(* IEC 61131-3 sources: daoli-st-library/DL_Device (part 31) *)

(* ---- FB_DL_SlurryLevelBank.st ---- *)
(*
  FB_DL_SlurryLevelBank  —  多罐浆料液位开关组（fail-safe 方向解释 / 质量字仲裁 / 开关相反归因）/ Slurry level switch bank
  分类 Category : DL_Device
  码位 Code     : 16#03_2_0E
  版本 Version  : 1.0.0
  来源 Source   : t2-8-isa182 — IEC 61131-3 标准语义的道莅防御性实现
  溯源 Origin   : ISA-18.2 报警管理公开语义借鉴（报警与故障分离、状态归因），clean-room 实现，未复制源码行
  功能 Function : 1) 逐罐读取高位/低位点式开关、质量字（0~3，0 = OK）与组态 fail-safe 方向；
                  2) 按 fail-safe 方向解释「液位 vs 断线」：LOW 型（eLow）断线时读数表现为高位，
                     HIGH 型（eHigh）断线时读数表现为低位——两类方向各自反推，绝不套用同一公式；
                  3) 质量字非 OK 判 abSensorFault，并以**安全侧**值参与联锁（保守取值：保护泵的取「低」，
                     保护溢流的取「高」，即一律认报警成立），信息级 011E 记录替代生效；
                  4) 同一罐高低位同时为真判「开关相反」故障 022E（3 罐 × 2 型共 6 组向量逐条推演，见验收向量）；
                  5) 输出严格区分「越限（工艺）」与「传感器故障（仪表）」两类：越限只置 abLevelAlarm 与信息级 010E，
                     传感器故障置 abSensorFault 与故障级 021E 并置 bError（R190 归因唯一）。
  边界 Boundary : ① uBankSize = 0 或 > DL_BANK_MAX 判组态错 020E，**直接返回不进入循环**（防数组越界，R28-2）；
                     高位/低位/质量字/方向四个数组声明长度一律 DL_BANK_MAX，长度不等在编译期即被拦截，
                     运行期再以 uBankSize 做上界闸（双保险）；
                  ② 质量字不在 0~3 域内判组态错（质量字编码越界，无法解释），不按 OK 处理；
                  ③ fail-safe 方向枚举落 ELSE（非法方向）按「最保守」处理：高低两位都认报警，并置 020E；
                  ④ 解除式自证：_bFault 清除 = rtReset.Q（引脚可满足）；022E 另可由「该罐高低位不再同时为真」
                     按码专清（R188 可达清除边，不依赖人工复位掩盖真实接线错误）；
                  ⑤ nFaultCount 为 INT，逐罐故障计数后钳制到 DL_BANK_MAX（不溢出、不回绕）；
                  ⑥ 越限（010E）为信息级，**永不置 bError**（R187③ / R45 配对纪律）。
  依赖 Depends  : 仅 Standard.library（TON / R_TRIG / ABS / MIN / MAX），零外部组件依赖
  同拍双窗配比  : tQualityDb（质量字去抖）与心跳窗 DL_HEART_WINDOW 不同源；配比约束
                  tQualityDb <= DL_HEART_WINDOW，保证去抖窗内至少一次判活（R100）

  码表 Error codes（本件格 03_2_0E，子码步进 +0x10）:
    16#0003_020E 故障级：组态非法（uBankSize = 0 或越上限 / 质量字越 0~3 域 / fail-safe 方向非法）
    16#0003_021E 故障级：传感器故障（质量字非 OK，已用安全侧值参与联锁）
    16#0003_022E 故障级：开关相反（同一罐高低位同时为真，接线或组态错误）
    16#0003_023E 故障级：状态机落 ELSE 兜底（非法相位 ID）
    16#0003_010E 信息级：液位越限（工艺告警，不置 bError）
    16#0003_011E 信息级：断线安全侧替代已生效（保守取值，不置 bError）

  修订历史 Revision :
    2026-11-18  v1.0.0  R37 首版
*)

TYPE E_DL_FailSafeDir :
(
    eLow  := 0,   // 低液位型：液位低时开关动作；断线时读数浮为「高位」/ Low-level type, a broken wire reads as high
    eHigh := 10   // 高液位型：液位高时开关动作；断线时读数浮为「低位」/ High-level type, a broken wire reads as low
);
END_TYPE

TYPE E_DL_LevelBankState :
(
    eIdle  := 0,   // 空闲：未使能，输出全部复位 / Idle, all outputs cleared while disabled
    eRun   := 10,  // 运行：逐罐评估 / Running, per-tank evaluation
    eFault := 90   // 故障：组态非法锁定 / Fault, illegal configuration latched
);
END_TYPE

FUNCTION_BLOCK FB_DL_SlurryLevelBank
VAR_INPUT
    bEnable        : BOOL := FALSE;                       // 总使能，FALSE 时输出全复位 / Master enable, low level clears the outputs
    bReset         : BOOL := FALSE;                       // 复位，上升沿清故障锁存 / Reset, rising edge clears the latch
    uBankSize      : UINT := 3;                           // 罐组实际罐数 [个]，域 1~DL_BANK_MAX / Number of tanks in use
    abLevelHigh    : ARRAY[0..7] OF BOOL;                 // 高位开关原始输入 [BOOL/罐] / Raw high-level switch inputs
    abLevelLow     : ARRAY[0..7] OF BOOL;                 // 低位开关原始输入 [BOOL/罐] / Raw low-level switch inputs
    anSensorQuality : ARRAY[0..7] OF INT;                 // 传感器质量字 [0~3，0 = OK] / Sensor quality word, zero means OK
    aeFailSafeDir  : ARRAY[0..7] OF E_DL_FailSafeDir;     // 每罐 fail-safe 方向组态 [枚举/罐] / Per-tank fail-safe direction
    tQualityDb     : TIME := T#500MS;                     // 质量字去抖窗 [ms]，域 > 0 / Quality debounce window [ms]
END_VAR
VAR_OUTPUT
    abLevelAlarm   : ARRAY[0..7] OF BOOL;                 // 逐罐液位越限报警 [BOOL/罐] / Per-tank level alarm
    abSensorFault  : ARRAY[0..7] OF BOOL;                 // 逐罐传感器故障 [BOOL/罐] / Per-tank sensor fault
    nFaultCount    : INT;                                 // 故障罐数 [个] / Number of faulty tanks
    bBankAlarm     : BOOL;                                // 罐组总报警（越限或故障任一）/ Bank aggregate alarm
    bValid         : BOOL;                                // 判据可用标志 / Criteria usable
    bError         : BOOL;                                // 故障标志，派生自锁存 / Fault flag derived from the latch
    nErrId         : UDINT;                               // 事件码，0 = 无事件 / Event code, 0 = no event
    eStateOut      : E_DL_LevelBankState;                 // 状态出口，段尾单点映射 / State outlet, mapped at the tail
END_VAR
VAR
    tonQuality   : TON;                                   // 质量故障去抖窗，每拍无条件调用 / Quality fault debounce, called unconditionally
    tonHeart     : TON;                                   // 周期心跳窗，自复位 / Periodic heartbeat window, self-resetting
    rtReset      : R_TRIG;                                // 复位上升沿 / Reset rising edge
    _eState      : E_DL_LevelBankState := E_DL_LevelBankState.eIdle;  // 内部相位（CASE 唯一写入目标）/ Internal phase
    _uFault      : UDINT;                                 // 故障码锁存 / Latched fault code
    _uInfo       : UDINT;                                 // 信息码，每拍重算 / Information code, recomputed per scan
    _bFault      : BOOL;                                  // 故障锁存位 / Latched fault bit
    _bCfgBad     : BOOL;                                  // 组态非法聚合 / Configuration invalid aggregate
    _bAnySensFault : BOOL;                                // 任一罐传感器故障 / Any sensor fault present
    _bAnyOpposite  : BOOL;                                // 任一罐高低位相反 / Any opposite-switch condition
    _bAnyLevelAlarm : BOOL;                               // 任一罐液位越限 / Any level alarm present
    _bSafeSubst  : BOOL;                                  // 本拍发生安全侧替代 / A safe-side substitution happened
    _bOppClear   : BOOL;                                  // 相反故障已全部消失 / All opposite conditions cleared
    _bHeartBrk   : BOOL := TRUE;                          // 心跳窗断输入一拍 / One-scan heartbeat break
    _bQualBrk    : BOOL := TRUE;                          // 质量去抖断输入一拍 / One-scan quality break
    _nIdx        : INT;                                   // 循环索引 [索引] / Loop index
    _nFaultAcc   : INT;                                   // 故障罐数保持量 [个] / Held faulty-tank count
    _bHighEff    : BOOL;                                  // 高位开关的解释后值（含安全侧替代）/ Effective high-level value
    _bLowEff     : BOOL;                                  // 低位开关的解释后值（含安全侧替代）/ Effective low-level value
    _bOpposite   : BOOL;                                  // 本罐高低位同时为真 / Both switches true in this tank
    _bQualBad    : BOOL;                                  // 本罐质量字非 OK / Quality word not OK in this tank
    _bDirBad     : BOOL;                                  // 本罐方向枚举非法 / Illegal direction enumeration in this tank
END_VAR
VAR CONSTANT
    DL_BANK_MAX   : INT := 8;          // 数组声明长度 [个]，四数组同长 / Declared array length, identical for all four arrays
    DL_QUAL_MAX   : INT := 3;          // 质量字最大值 [编码] / Maximum quality code
    DL_HEART_WINDOW : TIME := T#2S;    // 心跳观察窗 [ms]，自复位节拍 / Heartbeat window, self-resetting
END_VAR

(* —— 段 0：定时器与边缘检测无条件周期刷新（R182：调用语句不得置于 IF / CASE / FOR 内） —— *)
rtReset(CLK := bReset);                                          // 复位上升沿，每拍必调
tonHeart(IN := (NOT tonHeart.Q) AND (NOT _bHeartBrk), PT := DL_HEART_WINDOW);  // 心跳窗自复位
_bHeartBrk := FALSE;                                             // 断输入拍在调用后自清
tonQuality(IN := (_eState = E_DL_LevelBankState.eRun) AND _bAnySensFault AND (NOT _bQualBrk),
           PT := tQualityDb);                                    // 质量故障去抖（表达式入参）
_bQualBrk := FALSE;                                              // 断输入拍在调用后自清

(* —— 段 1：单拍量预清零（数组输出与保持量不入清单，R187①） —— *)
_uInfo        := 16#0000_0000;   // 信息码每拍重算
bError        := FALSE;          // 故障出口每拍重算，段 6 由锁存派生
bValid        := FALSE;          // 可用标志缺省 FALSE
bBankAlarm    := FALSE;          // 罐组总报警缺省 FALSE
_bCfgBad      := FALSE;          // 组态非法预清零
_bAnySensFault := FALSE;         // 传感器故障聚合预清零
_bAnyOpposite := FALSE;          // 相反故障聚合预清零
_bAnyLevelAlarm := FALSE;        // 越限聚合预清零
_bSafeSubst   := FALSE;          // 安全侧替代标志预清零
_bOppClear    := TRUE;           // 相反故障清空判定初值（循环内遇相反即置 FALSE）
_bDirBad      := FALSE;          // 方向非法预清零

(* —— 段 2：复位沿清锁存 + 按码专清（R188 双路径） —— *)
IF rtReset.Q THEN
    _bFault     := FALSE;            // 复位沿清锁存位
    _uFault     := 16#0000_0000;     // 复位沿清锁存码
    _nFaultAcc  := 0;                // 复位沿清故障罐数（重新统计）
END_IF

(* —— 段 3：组态域闸（循环之前完成，越界即返回不进入循环，R28-2） —— *)
IF (uBankSize = 0) OR (uBankSize > INT_TO_UINT(DL_BANK_MAX)) THEN
    _bCfgBad := TRUE;                // 罐数越界：0 或超数组声明长度
END_IF
IF TIME_TO_DINT(tQualityDb) <= 0 THEN
    _bCfgBad := TRUE;                // 去抖窗非法
END_IF
IF _bCfgBad THEN
    _uFault := 16#0003_020E;         // 故障级：组态非法
    _bFault := TRUE;                 // 锁存位置位（复位沿可清）
    bError  := TRUE;                 // 故障标志置位（R45 配对）
    _eState := E_DL_LevelBankState.eFault;  // 进故障相（不进入循环）
END_IF

(* —— 段 4：逐罐评估（仅运行相且组态合法时进入；循环上界由 uBankSize 钳制） —— *)
IF bEnable AND (_eState <> E_DL_LevelBankState.eFault) AND (NOT _bCfgBad) THEN
    _nFaultAcc := 0;                          // 故障罐数每拍重算（输出量，非台账）
    FOR _nIdx := 0 TO (UINT_TO_INT(uBankSize) - 1) DO
        (* 4.1 本罐假设值初始化：有效值先取原始值，随后按质量与方向修正 *)
        _bHighEff := abLevelHigh[_nIdx];       // 高位原始读数 [BOOL]
        _bLowEff  := abLevelLow[_nIdx];        // 低位原始读数 [BOOL]
        _bQualBad := (anSensorQuality[_nIdx] < 0) OR (anSensorQuality[_nIdx] > DL_QUAL_MAX) OR
                     (anSensorQuality[_nIdx] <> 0);            // 质量字非 OK（含越域：无法解释即判坏）
        IF (anSensorQuality[_nIdx] < 0) OR (anSensorQuality[_nIdx] > DL_QUAL_MAX) THEN
            _bCfgBad := TRUE;                  // 质量字越 0~3 域：组态/采集链错误
            _uFault := 16#0003_020E;           // 故障级：组态非法
            _bFault := TRUE;                   // 锁存
            bError  := TRUE;                   // 故障标志置位（R45 配对）
        END_IF
        IF _bQualBad THEN
            _bAnySensFault := TRUE;            // 传感器故障聚合
            abSensorFault[_nIdx] := TRUE;      // 逐罐故障输出
            _bSafeSubst := TRUE;               // 发生安全侧替代
            (* 4.2 fail-safe 方向解释：断线时 LOW 型读成「高位」，HIGH 型读成「低位」——
                   保守取值即两者都按「报警成立」处理（低液位保护泵、高液位保护溢流） *)
            IF aeFailSafeDir[_nIdx] = E_DL_FailSafeDir.eLow THEN
                _bHighEff := FALSE;            // LOW 型断线：原始高位读数是浮空假象，不予采信
                _bLowEff  := TRUE;             // 安全侧：认低液位（保护泵干转）
            ELSIF aeFailSafeDir[_nIdx] = E_DL_FailSafeDir.eHigh THEN
                _bHighEff := TRUE;             // 安全侧：认高液位（保护溢流）
                _bLowEff  := FALSE;            // HIGH 型断线：原始低位读数是浮空假象，不予采信
            ELSE
                _bDirBad := TRUE;              // 方向枚举非法：两位都认（最保守）
                _bHighEff := TRUE;
                _bLowEff  := TRUE;
                _uFault := 16#0003_020E;       // 故障级：组态非法（方向未组态）
                _bFault := TRUE;               // 锁存
                bError  := TRUE;               // 故障标志置位（R45 配对）
            END_IF
        ELSE
            abSensorFault[_nIdx] := FALSE;     // 质量 OK：清该罐传感器故障（按罐专清）
        END_IF
        (* 4.3 开关相反判据：同一罐高低位同时为真（物理上不可能，H 型与 L 型不可能同真） *)
        _bOpposite := _bHighEff AND _bLowEff;
        IF _bOpposite THEN
            _bAnyOpposite := TRUE;             // 相反故障聚合
            _bOppClear := FALSE;               // 相反条件仍在：禁止按码专清
            _uFault := 16#0003_022E;           // 故障级：开关相反
            _bFault := TRUE;                   // 锁存
            bError  := TRUE;                   // 故障标志置位（R45 配对）
        END_IF
        (* 4.4 越限判定：高低位任一为真即越限（信息级，不置 bError） *)
        IF _bHighEff OR _bLowEff THEN
            abLevelAlarm[_nIdx] := TRUE;       // 逐罐越限输出
            _bAnyLevelAlarm := TRUE;           // 越限聚合
        ELSE
            abLevelAlarm[_nIdx] := FALSE;      // 本罐无越限：按罐清零
        END_IF
        (* 4.5 故障罐数累计：传感器故障 + 开关相反各计一次（越限不计入故障数） *)
        IF abSensorFault[_nIdx] OR _bOpposite THEN
            IF _nFaultAcc < DL_BANK_MAX THEN
                _nFaultAcc := _nFaultAcc + 1;  // 故障罐数 +1（钳制到声明长度，不溢出）
            END_IF
        END_IF
    END_FOR
    (* 4.6 未使用的罐位输出清零（上界之外不得残留旧值） *)
    FOR _nIdx := UINT_TO_INT(uBankSize) TO (DL_BANK_MAX - 1) DO
        abLevelAlarm[_nIdx]  := FALSE;         // 未用罐位：越限清零
        abSensorFault[_nIdx] := FALSE;         // 未用罐位：故障清零
    END_FOR
ELSE
    _nFaultAcc := 0;                           // 故障相/组态非法：不做评估，故障数为 0（不伪造）
    FOR _nIdx := 0 TO (DL_BANK_MAX - 1) DO
        abLevelAlarm[_nIdx]  := FALSE;         // 全清：越限输出
        abSensorFault[_nIdx] := TRUE;          // 全置：故障相时无法判读，按不可信上报
    END_FOR
END_IF

(* —— 段 5：相位机（只做迁移；输出映射在段 7，CASE 内不写输出枚举，N2） —— *)
CASE _eState OF
E_DL_LevelBankState.eIdle:
    _nFaultAcc := 0;                           // 空闲：不做评估，故障罐数归零
    IF bEnable AND (NOT _bCfgBad) AND (NOT _bFault) THEN
        _eState := E_DL_LevelBankState.eRun;   // 使能且组态合法：进运行相
    END_IF
E_DL_LevelBankState.eRun:
    IF NOT bEnable THEN
        _eState := E_DL_LevelBankState.eIdle;  // 失能：回空闲（输出在段 7 单点清零）
    END_IF
E_DL_LevelBankState.eFault:
    IF (NOT _bFault) AND (NOT _bCfgBad) AND bEnable THEN
        _eState := E_DL_LevelBankState.eRun;   // 锁存已清且组态合法：回运行相
    END_IF
ELSE
    _uFault := 16#0003_023E;                   // 故障级：相位 ID 越界（枚举兜底）
    _bFault := TRUE;                           // 锁存
    bError  := TRUE;                           // 故障标志置位（R45 配对）
    _eState := E_DL_LevelBankState.eFault;     // 强制回故障相
END_CASE

(* 段 5B｜按码专清（依赖段 4 的逐罐结果，故必须置于评估之后，R188 可达清除边） *)
IF (_uFault = 16#0003_022E) AND _bOppClear THEN
    _uFault := 16#0000_0000;                   // 相反条件全部消失 → 该码可解
    _bFault := FALSE;                          // 锁存位同步清
END_IF
IF (_uFault = 16#0003_021E) AND (NOT _bAnySensFault) AND (NOT _bCfgBad) THEN
    _uFault := 16#0000_0000;                   // 质量字全部恢复 OK → 传感器故障码可解
    _bFault := FALSE;                          // 锁存位同步清
END_IF

(* —— 段 6：信息码与故障码优先级链（越限永不置 bError；每个 bError 源均有码，R45） —— *)
IF _bAnySensFault AND _bSafeSubst THEN
    _uInfo := 16#0003_011E;                    // 信息级：断线安全侧替代已生效
ELSIF _bAnyLevelAlarm THEN
    _uInfo := 16#0003_010E;                    // 信息级：液位越限（工艺告警）
END_IF
IF _bCfgBad THEN
    _uFault := 16#0003_020E;                   // 组态非法优先上报（其余码不得掩盖组态根因）
    _bFault := TRUE;                           // 锁存
    bError  := TRUE;                           // 故障标志置位
ELSIF _bAnyOpposite THEN
    _uFault := 16#0003_022E;                   // 开关相反优先于传感器故障上报（接线错根因）
    _bFault := TRUE;                           // 锁存
    bError  := TRUE;                           // 故障标志置位
ELSIF _bAnySensFault AND tonQuality.Q THEN
    _uFault := 16#0003_021E;                   // 传感器故障：去抖窗满才上报（防瞬时质量抖动）
    _bFault := TRUE;                           // 锁存
    bError  := TRUE;                           // 故障标志置位
END_IF

(* —— 段 7：出口单点映射（名实同源；锁存码回放，禁同拍抹除） —— *)
IF _eState = E_DL_LevelBankState.eIdle THEN
    FOR _nIdx := 0 TO (DL_BANK_MAX - 1) DO
        abLevelAlarm[_nIdx]  := FALSE;         // 空闲：越限输出清零
        abSensorFault[_nIdx] := FALSE;         // 空闲：故障输出清零
    END_FOR
END_IF
nFaultCount := _nFaultAcc;                     // 故障罐数出口
bBankAlarm  := _bAnyLevelAlarm OR _bAnyOpposite OR _bAnySensFault OR _bFault;  // 罐组总报警
eStateOut   := _eState;                        // 状态出口
IF _bFault THEN
    nErrId := _uFault;                         // 故障锁存码回放（不在故障相按当下输入重推）
    bError := TRUE;                            // 故障出口派生自锁存
ELSE
    nErrId := _uInfo;                          // 信息码
END_IF
bValid := bEnable AND (NOT _bFault) AND (NOT _bCfgBad);  // 判据可用

END_FUNCTION_BLOCK

(* ---- FB_DL_SlurryStirrerCtrl.st ---- *)
(*==============================================================================
 * 组件名称 (Component)  : FB_DL_SlurryStirrerCtrl
 * 所属子库 (Sublibrary) : DL_Device
 * 前缀     (Prefix)     : FB_DL_
 * 当前版本 (Version)    : 1.0.0
 * 兼容性   (Platform)   : CODESYS 3.5 / TwinCAT 3 / 汇川 InoProShop / Schneider
 *                         Machine Expert；纯 IEC 61131-3（第 3 版），
 *                         仅依赖标准库 TON / R_TRIG / ABS / MAX / MIN，零厂商方言
 * 作者     (Author)     : 道莅代码库 · PLC编程专家（R31）
 * 开源溯源 (Origin)     : 浆料搅拌双电机同步控制公开工艺语义（行业池），
 *                         道莅 clean-room 防御性实现，未复制任何外部源码行
 * 功能描述 (Function)   : 浆料搅拌双电机同步件。双电机主从同启（启差不超过
 *                         tSync 防涌流）；同步监视为两机扭矩偏差百分数超
 *                         fSyncTol 持续 tConf 即摘从机降级；单机扭矩超
 *                         fTrqMax 持续 tConf 停该机锁故障。扭矩非有限按
 *                         传感器失效摘除该机，不猜值。等级到健康映射写死
 *                         本头注释。粘度趋势判据依赖库内 FB_DL_Differentiator
 *                         （引脚注入消费，不内联），见依赖表。
 * 依赖表   (Depends)    : E_DL_Ne107Status（属主 I_DL_DeviceHealth.st，只引用
 *                         不重声明）；FB_DL_Differentiator（上层粘度趋势
 *                         判据注入消费，本件本体不调用）。
 * 健康映射 (Health map) : eFailure = 扭矩超限锁故障；eMaintenanceReq = 同步
 *                         失稳摘从机降级；eOutOfSpec = 传感器失效摘除；
 *                         eCheckFunction = 启动暂态（主从启差期间）；eOk = 正常。
 * 码位     (Codes)      : 16#0003_03F7 信息级：传感器失效摘除、参数钳位、
 *                                      扭矩监视禁用（不置 bError）
 *                         16#0003_03F8 故障级：单机扭矩超限（锁存）
 *                         16#0003_03F9 故障级：同步失稳（锁存）
 *                         16#0003_03FA 故障级：状态非法（ELSE 兜底，锁存）
 *                         16#0003_03FB 保留未启用（码表与实现对齐，不虚声明）
 * 边界防错 (Boundary)   : 1 扭矩非有限（x<>x 自反判加幅值界）摘该机不猜值；
 *                         2 均值防除零取 max(均值, 1.0E-6)；
 *                         3 TON/R_TRIG 实例每拍无条件刷新；
 *                         4 CASE 带 ELSE 锁故障兜底；
 *                         5 故障锁存可达解除路径：bRun 撤除回待机清码；
 *                         6 fSyncTol 非正钳 1.0；fTrqMax 非正禁用超限监视并
 *                           记信息码（禁用留档，不静默）。
 * 修订历史 (Revision)   : 2026-11-18 v1.0.0 首版入库（R31 · 阶段三 · 序 10）
 *==============================================================================*)

(*------------------------------------------------------------------------------
 * 枚举: E_DL_StirState（归属本功能块，同文件发布，全库唯一属主）
 *----------------------------------------------------------------------------*)
TYPE E_DL_StirState :
(
    eIdle     := 0,    // 待机：双机停 / Idle, both motors stopped
    eStart1   := 10,   // 主机启动态：仅主机得电 / Main-start state, main motor only
    eRun      := 20,   // 双机运行态：主从同步 / Run state, both motors synchronized
    eDegrade  := 30,   // 降级态：从机已摘除 / Degraded state, follower removed
    eFault    := 99    // 故障态：锁存等待撤运行 / Fault state, latched until run dropped
);
END_TYPE

(*==============================================================================
 * 功能块: FB_DL_SlurryStirrerCtrl
 * 调用约定: 每个扫描周期无条件调用一次；扭矩信号经引脚注入。
 *==============================================================================*)
FUNCTION_BLOCK FB_DL_SlurryStirrerCtrl
VAR_INPUT
    bRun     : BOOL := FALSE;         // 运行指令（电平）/ Run command, level active
    fTrq1    : REAL := 0.0;           // 电机 1 扭矩 [牛米] / Motor 1 torque [Nm]
    fTrq2    : REAL := 0.0;           // 电机 2 扭矩 [牛米] / Motor 2 torque [Nm]
    fTrqMax  : REAL := 50.0;          // 单机扭矩上限 [牛米]，非正禁用监视 / Per-motor torque limit [Nm], non-positive disables monitor
    fSyncTol : REAL := 10.0;          // 同步偏差容差 [百分数] / Sync deviation tolerance [%]
    tConf    : TIME := T#2S;          // 判级确认时长 [毫秒] / Judgement confirm duration [ms]
    tSync    : TIME := T#1S;          // 主从启差上限 [毫秒] / Start stagger limit [ms]
END_VAR
VAR_OUTPUT
    bStart1  : BOOL;                  // 电机 1 启动指令 / Motor 1 start command
    bStart2  : BOOL;                  // 电机 2 启动指令 / Motor 2 start command
    bSyncOk  : BOOL;                  // 同步合格标志 / Synchronization OK flag
    eHealth  : E_DL_Ne107Status;      // 健康出口（引用库内枚举，只引用不重声明）/ Health output, library enum referenced only
    bError   : BOOL;                  // 故障标志，与故障级码配对（R45）/ Fault flag paired with fault codes
    uErrorId : UDINT;                 // 错误码，0 = 无错 / Error code, 0 = none
END_VAR
VAR
    rTrigRun : R_TRIG;                // 运行沿检测，每拍无条件刷新 / Run edge detector, refreshed every scan
    tonStag  : TON;                   // 主从启差定时器，每拍无条件刷新 / Start stagger timer, refreshed every scan
    tonSync  : TON;                   // 同步失稳确认定时器，每拍无条件刷新 / Sync instability timer, refreshed every scan
    tonTrq   : TON;                   // 扭矩超限确认定时器，每拍无条件刷新 / Torque overlimit timer, refreshed every scan
    eState   : E_DL_StirState;        // 内部状态机 / Internal state machine
    bSen1Ok  : BOOL;                  // 电机 1 传感器有效 / Motor 1 sensor valid
    bSen2Ok  : BOOL;                  // 电机 2 传感器有效 / Motor 2 sensor valid
    bSenBad  : BOOL;                  // 任一传感器失效 / Any sensor failed
    bDevNow  : BOOL;                  // 本拍同步偏差超限 / Sync deviation out of band this scan
    bOv1     : BOOL;                  // 电机 1 扭矩超限 / Motor 1 torque overlimit
    bOv2     : BOOL;                  // 电机 2 扭矩超限 / Motor 2 torque overlimit
    bOvNow   : BOOL;                  // 本拍任一机超限 / Any overlimit this scan
    fTolEff  : REAL;                  // 钳位后生效容差 [百分数] / Effective clamped tolerance [%]
    fDevPct  : REAL;                  // 扭矩偏差百分数 [%] / Torque deviation percent [%]
    fMean    : REAL;                  // 双机扭矩均值防除零基准 [牛米] / Torque mean with divide guard [Nm]
    bTrqMonOn: BOOL;                  // 超限监视使能（上限合法）/ Overlimit monitor enabled
    uCodeLatch: UDINT;                // 故障级锁存码 / Latched fault code
    bInfoTrq : BOOL;                  // 本拍参数/监视禁用信息 / Parameter or monitor info this scan
END_VAR
VAR CONSTANT
    DL_SSC_FIN   : REAL := 1.0E30;    // REAL 有限幅值判界 / REAL finiteness magnitude bound
    DL_SSC_EPS   : REAL := 1.0E-6;    // 均值防除零容差 [牛米] / Mean divide-guard tolerance [Nm]
    DL_SSC_TOLMIN: REAL := 1.0;       // 同步容差钳位下限 [百分数] / Tolerance clamp floor [%]
    DL_SSC_PCT   : REAL := 100.0;     // 百分数换算系数 / Percent conversion factor
END_VAR

// ---- 段 1｜边沿与定时器实例无条件周期刷新（红线：禁入条件分支）----------------
rTrigRun(CLK := bRun);                                // 运行沿检测 / Run edge detection
tonStag(IN := (eState = eStart1), PT := tSync);       // 启差计时按态断输入 / Stagger timing input per state
tonSync(IN := bDevNow, PT := tConf);                  // 失稳确认无条件计时 / Instability timing unconditionally
tonTrq(IN := bOvNow, PT := tConf);                    // 超限确认无条件计时 / Overlimit timing unconditionally

// ---- 段 2｜传感器有效性与参数钳位 ----------------------------------------------
bSen1Ok := (fTrq1 = fTrq1) AND (ABS(fTrq1) < DL_SSC_FIN); // 电机 1 扭矩有限 / Motor 1 torque finite
bSen2Ok := (fTrq2 = fTrq2) AND (ABS(fTrq2) < DL_SSC_FIN); // 电机 2 扭矩有限 / Motor 2 torque finite
bSenBad := (NOT bSen1Ok) OR (NOT bSen2Ok);            // 任一失效 / Any sensor failed
fTolEff := fSyncTol;                                  // 容差原值 / Tolerance as-is
bInfoTrq := FALSE;                                    // 信息标志先清 / Clear info flag
IF fTolEff <= 0.0 THEN
    fTolEff := DL_SSC_TOLMIN;                         // 非正容差钳下限 / Clamp non-positive tolerance
    bInfoTrq := TRUE;                                 // 记参数钳位 / Record parameter clamp
END_IF
bTrqMonOn := (fTrqMax > 0.0) AND (fTrqMax < DL_SSC_FIN); // 上限合法才使能监视 / Monitor only with legal limit
IF NOT bTrqMonOn THEN
    bInfoTrq := TRUE;                                 // 监视禁用记信息码 / Monitor disabled records info
END_IF

// ---- 段 3｜同步偏差与超限判据（均值防除零）--------------------------------------
IF bSen1Ok AND bSen2Ok THEN
    fMean := MAX(0.5 * (ABS(fTrq1) + ABS(fTrq2)), DL_SSC_EPS); // 均值防除零 / Mean with divide guard
    fDevPct := ABS(fTrq1 - fTrq2) / fMean * DL_SSC_PCT;        // 偏差百分数 / Deviation percent
    bDevNow := fDevPct > fTolEff;                              // 本拍超差 / Out of band this scan
    bOv1 := bTrqMonOn AND (fTrq1 > fTrqMax);                   // 电机 1 超限判定 / Motor 1 overlimit
    bOv2 := bTrqMonOn AND (fTrq2 > fTrqMax);                   // 电机 2 超限判定 / Motor 2 overlimit
ELSE
    fDevPct := 0.0;                                            // 异常路径确定值 / Deterministic fallback
    bDevNow := FALSE;                                          // 传感器失效不判同步 / No sync judge with bad sensor
    bOv1 := FALSE;                                             // 失效机不判超限 / No overlimit judge
    bOv2 := FALSE;                                             // 失效机不判超限 / No overlimit judge
END_IF
bOvNow := bOv1 OR bOv2;                                        // 任一超限 / Any overlimit

// ---- 段 4｜状态机（CASE 带 ELSE 锁故障兜底）--------------------------------------
CASE eState OF
    eIdle:
        bStart1 := FALSE;                             // 待机双机停 / Both stopped in idle
        bStart2 := FALSE;                             // 待机双机停 / Both stopped in idle
        IF rTrigRun.Q THEN
            eState := eStart1;                        // 运行沿进主机启动 / Run edge starts main motor
        END_IF
    eStart1:
        bStart1 := bRun;                              // 主机随运行指令 / Main follows run command
        bStart2 := FALSE;                             // 从机未得电 / Follower not powered
        IF NOT bRun THEN
            eState := eIdle;                          // 撤运行回待机 / Run drop returns to idle
        ELSIF tonStag.Q THEN
            eState := eRun;                           // 启差满双机运行 / Stagger elapsed, both run
        END_IF
    eRun:
        bStart1 := bRun AND bSen1Ok;                  // 主机指令带传感器门控 / Main gated by sensor
        bStart2 := bRun AND bSen2Ok AND (NOT tonSync.Q); // 从机失稳即摘除 / Follower removed on instability
        IF NOT bRun THEN
            eState := eIdle;                          // 撤运行回待机 / Run drop returns to idle
        ELSIF tonTrq.Q THEN
            eState := eFault;                         // 超限确认锁故障 / Overlimit confirmed, fault
            uCodeLatch := 16#0003_03F8;               // 码位：扭矩超限 / Code: torque overlimit
        ELSIF tonSync.Q THEN
            eState := eDegrade;                       // 同步失稳摘从机降级 / Sync lost, degrade
            uCodeLatch := 16#0003_03F9;               // 码位：同步失稳 / Code: sync instability
        END_IF
    eDegrade:
        bStart1 := bRun AND bSen1Ok;                  // 降级态仅主机 / Only main in degraded
        bStart2 := FALSE;                             // 从机保持摘除 / Follower stays removed
        IF NOT bRun THEN
            eState := eIdle;                          // 可达解除：撤运行回待机清码 / Reachable release: run drop
            uCodeLatch := 16#0000_0000;               // 清锁存码 / Clear latched code
        END_IF
    eFault:
        bStart1 := FALSE;                             // 故障停主机（该机）/ Main stopped in fault
        bStart2 := FALSE;                             // 故障停从机 / Follower stopped in fault
        IF NOT bRun THEN
            eState := eIdle;                          // 可达解除：撤运行回待机 / Reachable release: run drop
            uCodeLatch := 16#0000_0000;               // 清锁存码 / Clear latched code
        END_IF
    ELSE
        eState := eFault;                             // 非法状态兜底 / Illegal state fallback
        uCodeLatch := 16#0003_03FA;                   // 码位：状态非法 / Code: illegal state
END_CASE

// ---- 段 5｜同步合格与健康出口装配（映射写死头注释）------------------------------
bSyncOk := (eState = eRun) AND (NOT bDevNow) AND (NOT bSenBad) AND (NOT bOvNow); // 同步合格 / Sync OK
IF eState = eFault THEN
    eHealth := eFailure;                              // 扭矩超限锁故障 / Torque overlimit failure
ELSIF eState = eDegrade THEN
    eHealth := eMaintenanceReq;                       // 失稳降级 / Degraded maintenance
ELSIF bSenBad THEN
    eHealth := eOutOfSpec;                            // 传感器失效摘除 / Sensor failure out-of-spec
ELSIF eState = eStart1 THEN
    eHealth := eCheckFunction;                        // 启动暂态 / Starting transient
ELSIF (eState = eRun) OR (eState = eIdle) THEN
    eHealth := eOk;                                   // 正常 / Normal
ELSE
    eHealth := eUnknown;                              // 兜底未知 / Fallback unknown
END_IF

// ---- 段 6｜错误码装配：故障锁存回放优先，信息级居次 ------------------------------
IF eState = eFault THEN
    bError   := TRUE;                                 // 故障标志配对（R45）/ Fault flag paired
    uErrorId := uCodeLatch;                           // 故障码锁存回放 / Latched fault code replayed
ELSIF bSenBad OR bInfoTrq THEN
    bError   := FALSE;                                // 信息级不置故障 / Info never sets fault
    uErrorId := 16#0003_03F7;                         // 信息级：失效/钳位/禁用 / Info: sensor or parameter
ELSE
    bError   := FALSE;                                // 无错清标志 / Clear fault flag
    uErrorId := 16#0000_0000;                         // 无码 / No code
END_IF
END_FUNCTION_BLOCK

(* ---- FB_DL_SoakPitTemperatureCtrl.st ---- *)
(*
  Component : FB_DL_SoakPitTemperatureCtrl
  Category  : DL_Device
  Type      : FB
  Complexity: C2
  VERSION   : v1.0.0
  功能      : 坑式炉均热控制：设定-实测偏差带内做简化 PI（比例 + 积分限幅）输出加热百分比，偏差带内持续驻留到时报均热完成。
  开源溯源  : 道莅原创 clean-room 自研（无外部代码引用）｜License: MIT
  边界条件  : ① 偏差带、采样周期、输出上限须 > 1e-9，否则判组态非法并锁存故障；
              ② 积分项做 0~输出上限双侧限幅（抗饱和），使能撤销时积分清零；
              ③ 均热完成位为锁存置位，仅在使能撤销或复位沿清除。
*)
FUNCTION_BLOCK FB_DL_SoakPitTemperatureCtrl
VAR_INPUT
    bEnable    : BOOL;   (* 使能电平 [-] Enable level *)
    bReset     : BOOL;   (* 复位上升沿，清完成位与故障 [-] Reset edge *)
    fSetC      : REAL;   (* 均热温度设定 [°C] Soaking temperature setpoint *)
    fActC      : REAL;   (* 炉膛实测温度 [°C] Measured furnace temperature *)
    fKp        : REAL;   (* 比例增益 [%/K] Proportional gain *)
    fKi        : REAL;   (* 积分增益 [%/(K·s)] Integral gain *)
    fOutMaxPct : REAL;   (* 加热输出上限 [%] Heater output upper limit *)
    fBandC     : REAL;   (* 均热偏差带半宽 [K] Soaking band half width *)
    tSample    : TIME;   (* PI 采样周期 [ms] PI sampling period *)
    tSoakDur   : TIME;   (* 均热驻留时长 [ms] Soaking dwell time *)
END_VAR
VAR_OUTPUT
    fOutPct    : REAL;   (* 加热输出百分比 [%] Heater output percent *)
    fErrC      : REAL;   (* 当前温度偏差 [K] Current temperature error *)
    bInBand    : BOOL;   (* 偏差带内标志 [-] Within band flag *)
    bSoakDone  : BOOL;   (* 均热完成（锁存） [-] Soaking done latched *)
    bError     : BOOL;   (* 故障锁存标志 [-] Fault latch flag *)
    uErrId     : UDINT;  (* 事件码，0 = 无事件 [-] Event code *)
END_VAR
VAR
    rtReset  : R_TRIG;   (* 复位沿实例，每拍无条件刷新 / Reset edge *)
    tonSample: TON;      (* 采样节拍（自复位错峰） / Sampling tick self-reset *)
    tonSoak  : TON;      (* 均热驻留计时（独立实例） / Soaking dwell timer *)
    _fInteg  : REAL;     (* 积分累计量 [%] Integral accumulator *)
    _bDone   : BOOL;     (* 均热完成锁存位（锁存量） / Latched done bit *)
    _bFault  : BOOL;     (* 故障锁存位（锁存量） / Latched fault bit *)
    _uFault  : UDINT;    (* 故障码锁存（锁存量） / Latched fault code *)
    _bCfgBad : BOOL;     (* 组态非法当拍量 [-] Config illegal flag *)
    _bNonFin : BOOL;     (* 输入非有限当拍量 [-] Non-finite input flag *)
    fDt      : REAL;     (* 采样周期秒值 [s] Sampling period in seconds *)
END_VAR
VAR CONSTANT
    DL_EPS     : REAL := 1.0E-9;    (* 除零判定容差 [无量纲] Divide-by-zero tolerance *)
    DL_MS_PER_S: REAL := 1000.0;    (* 毫秒转秒换算系数 [ms/s] Milliseconds per second *)
    DL_ZERO    : REAL := 0.0;       (* 零常量 [无量纲] Zero constant *)
END_VAR

(* —— 段 1｜每拍量预清零（锁存量 _bDone/_bFault/_uFault/_fInteg 不入清单） —— *)
uErrId := 16#0000_0000;
_bCfgBad := FALSE;
_bNonFin := FALSE;

(* —— 段 2｜非有限拦截与组态闸（覆盖采样周期、偏差带、输出上限、增益） —— *)
IF (fActC <> fActC) OR ((fActC - fActC) <> 0.0)
   OR (fSetC <> fSetC) OR ((fSetC - fSetC) <> 0.0)
   OR (fKp <> fKp) OR ((fKp - fKp) <> 0.0)
   OR (fKi <> fKi) OR ((fKi - fKi) <> 0.0)
   OR (fOutMaxPct <> fOutMaxPct) OR ((fOutMaxPct - fOutMaxPct) <> 0.0)
   OR (fBandC <> fBandC) OR ((fBandC - fBandC) <> 0.0) THEN
    _bNonFin := TRUE;
END_IF
IF (fBandC <= DL_EPS) OR (fOutMaxPct <= DL_EPS) OR (fKp < DL_ZERO) OR (fKi < DL_ZERO)
   OR (tSample = T#0S) OR (tSoakDur = T#0S) THEN
    _bCfgBad := TRUE;
END_IF
IF _bCfgBad AND (NOT _bFault) THEN
    _bFault := TRUE;
    _uFault := 16#0022_0001;              (* 故障级：组态非法 / Fault code bad config *)
END_IF
IF _bNonFin AND (NOT _bFault) THEN
    _bFault := TRUE;
    _uFault := 16#0022_0002;              (* 故障级：温度反馈非有限 / Non-finite temperature *)
END_IF

(* —— 段 3｜偏差与带内判定（本拍值，先于定时器使用） —— *)
fErrC := fSetC - fActC;                   (* 偏差 = 设定 - 实测 [K] *)
IF fErrC < DL_ZERO THEN
    bInBand := (-fErrC) <= fBandC;        (* 负偏差取绝对值比较 [K] / Absolute compare *)
ELSE
    bInBand := fErrC <= fBandC;           (* 正偏差直接比较 [K] / Direct compare *)
END_IF

(* —— 段 4｜沿与定时器每拍无条件刷新（tonSample 自复位错峰，禁靠外部沿清零） —— *)
rtReset  (CLK := bReset);
tonSample(IN := NOT tonSample.Q, PT := tSample);
tonSoak  (IN := bInBand AND bEnable AND (NOT _bFault), PT := tSoakDur);

(* —— 段 5｜复位沿：清完成位、积分与故障（唯一解除路径） —— *)
IF rtReset.Q THEN
    _bFault := FALSE;
    _uFault := 16#0000_0000;
    _bDone := FALSE;
    _fInteg := DL_ZERO;
END_IF

(* —— 段 6｜简化 PI：每个采样节拍做一次积分，积分与输出双侧限幅（抗饱和） —— *)
fDt := TIME_TO_REAL(tSample) / DL_MS_PER_S;
IF tonSample.Q THEN
    IF fDt > DL_EPS THEN
        _fInteg := _fInteg + fKi * fErrC * fDt;
    END_IF
    IF _fInteg > fOutMaxPct THEN
        _fInteg := fOutMaxPct;            (* 积分上限限幅 [%] / Integral upper clamp *)
    ELSIF _fInteg < DL_ZERO THEN
        _fInteg := DL_ZERO;               (* 积分下限限幅 [%] / Integral lower clamp *)
    END_IF
END_IF
IF bEnable AND (NOT _bFault) THEN
    fOutPct := fKp * fErrC + _fInteg;
    IF fOutPct > fOutMaxPct THEN
        fOutPct := fOutMaxPct;            (* 输出上限限幅 [%] / Output upper clamp *)
    ELSIF fOutPct < DL_ZERO THEN
        fOutPct := DL_ZERO;               (* 输出下限限幅 [%] / Output lower clamp *)
    END_IF
ELSE
    fOutPct := DL_ZERO;                   (* 非使能：输出归零、积分复位 *)
    _fInteg := DL_ZERO;
    _bDone := FALSE;
END_IF

(* —— 段 7｜均热完成锁存：驻留到置位，只认复位沿或使能撤销 —— *)
IF tonSoak.Q THEN
    _bDone := TRUE;
END_IF

(* —— 段 8｜出口单点映射 —— *)
bSoakDone := _bDone;
bError := _bFault;
IF _bFault AND (_uFault <> 16#0000_0000) THEN
    uErrId := _uFault;                    (* 故障码锁存回放 / Latched fault replay *)
END_IF
END_FUNCTION_BLOCK

(* ---- FB_DL_SoftStarterDrive.st ---- *)
(*
  ==================================================================
  组件名 Component  : FB_DL_SoftStarterDrive
  分类   Category   : DL_Device
  复杂度 Complexity  : cx5
  版本   Version    : 1.0.1
  功能   Purpose    : 软启动器驱动封装。晶闸管斜坡启动（bCmdRun 端子）→ 斜坡
                      末投旁路接触器（bCmdBypass）→ 旁路反馈确认转运行；停
                      机双命令全断 + 旁路分断确认；斜坡窗 / 反馈确认窗 / 停
                      机确认窗三窗监视 + 启动超时保护 + 旁路提前吸合矛盾诊
                      断 + 过载锁存 + 重启抑制冷却。实现既有 I_DL_MotorDriver
                      接口，补齐 DOL / 星三角 / 软启 / 变频四启动家族。
  来源   Source     : t2-2-lbp（cmd / ind 分离范式）
  溯源   Origin     : IEC 61131-3 标准语义的道莅防御性实现；软启动器旁路投
                      切与反馈校验为行业公知工程语义，clean-room 自研实现，
                      未复制 LBP 或任何厂商私有库源码。
  平台   Platform   : 纯 IEC 61131-3（Standard.library: TON / R_TRIG，无私有库）
  接口实现 Implements : I_DL_MotorDriver（属主文件 DL_Device\I_DL_MotorDriver.st）。
                      R66 收窄清单：契约属性 eState / bRunning / bFault /
                      uErrorId / bRestartInhibit 仅以 PROPERTY GET 落地（本件
                      不在 VAR_OUTPUT 重复声明同名引脚）；方法 CmdStart /
                      CmdStop / CmdReset 签名一字不减，契约语义一字不减。
  平台枚举归属 Ownership : 内部状态映射 E_DL_MotorState（归属 I_DL_MotorDriver
                      同文件发布，本件只引用不重声明）。
  码位留痕 CodeSource : 实现 I_DL_MotorDriver 契约 uErrorId（接口文件声明段位
                      16#0003_xxxx），沿用族内既有派号段（FB_DL_DolMotor 已占
                      0201..020A），本件占用 0211..0217：故障级 0003_0211 旁路
                      反馈确认超时 / 0003_0212 运行中旁路反馈断开 / 0003_0213
                      停机旁路未分断 / 0003_0214 斜坡期旁路提前吸合 / 0003_0215
                      过载锁存 / 0003_0216 非法状态；信息级 0003_0217 重启抑制
                      期拒绝（只写 uErrorId 不进 bFault，0.2 公约）。锁存解除
                      路径 = bReset 上升沿（唯一路径，R188）。
  作者   Author     : 道莅代码库 · PLC 编程专家（R58）
  ------------------------------------------------------------------
  边界 Boundary     :
                      一 三窗配比约束（R100）：tFbWindow < tRampTime（旁路反
                         馈窗必须短于斜坡窗）且 tStopConfirm < tRestartInhibit
                         （停机确认短于冷却窗）；越域由调用方组态保证，本件
                         不做二次钳制；
                      二 停机双命令全断：bCmdRun 与 bCmdBypass 在停机 / 故障
                         / 过载相安全侧全断（R191 降级显式声明）；
                      三 过载全局监视优先级最高：斜坡 / 投旁路 / 运行相过载
                         立即锁存脱扣（R190 独立成因独立码）；
                      四 方法均为非阻塞单发，跨周期动作由 _bPend* 请求标志
                         交主体状态机消化（无 METHOD 内状态驻留）；
                      五 无全局变量、无外部变量声明、无物理地址寻址。
  修订记录 Revision  :
    2026-11-21  v1.0.0  R58 首版（批 2 · 序号 7）
    2026-11-21  v1.0.1  R59 返修轻①②：复位分支前置故障相位门（故障相复位只清锁存不迁相）；删 3 处 _ePhase 自赋值死语句
  ==================================================================
*)

TYPE E_DL_SsdPhase :
(
    eSsdIdle    := 0,  // 空闲：消化停止锁存，评估启动请求 / idle, absorbing the stop latch
    eSsdRamp    := 10, // 晶闸管斜坡：运行端子得电，旁路断开 / the thyristor ramp, the run terminal on, the bypass off
    eSsdByWait  := 20, // 投旁路：旁路命令得电，等反馈吸合确认 / the bypass engage, the command on, awaiting the feedback
    eSsdRun     := 30, // 旁路运行：反馈吸合确认带载 / the bypass running, feedback confirmed
    eSsdStop    := 40, // 停机过渡：双命令全断，等旁路分断确认 / the stopping transition, both commands off, awaiting the drop out
    eSsdTrip    := 50, // 过载脱扣锁存：仅复位且过载消失可清 / the overload trip latch
    eSsdFault   := 90  // 故障锁存：仅复位可清 / the latched fault
);
END_TYPE

FUNCTION_BLOCK FB_DL_SoftStarterDrive IMPLEMENTS I_DL_MotorDriver
VAR_INPUT
    bCmdStart       : BOOL;           // 启动指令，上升沿生效 [-] / the start command, rising edge effective
    bCmdStop        : BOOL;           // 停止指令，电平生效 [-] / the stop command, level effective
    bFbBypass       : BOOL := FALSE;  // 旁路接触器反馈，TRUE = 吸合 [-] / the bypass contactor feedback, true = picked up
    bOverload       : BOOL := FALSE;  // 过载保护信号，TRUE = 过载 [-] / the overload protection signal, true = overloaded
    bPermitStart    : BOOL := TRUE;   // 启动允许联锁，TRUE = 允许 [-] / the start permit interlock, true = allowed
    tRampTime       : TIME := T#10S;  // 晶闸管斜坡时长 [毫秒] / the thyristor ramp duration [millisecond]
    tFbWindow       : TIME := T#2S;   // 旁路反馈确认窗 [毫秒] / the bypass feedback confirm window [millisecond]
    tStopConfirm    : TIME := T#5S;   // 停机旁路分断确认窗 [毫秒] / the stop drop out confirm window [millisecond]
    tRestartInhibit : TIME := T#60S;  // 重启抑制冷却时长 [毫秒] / the restart inhibit cooling duration [millisecond]
    bReset          : BOOL;           // 故障复位，上升沿生效 [-] / the fault reset, rising edge effective
END_VAR
VAR_OUTPUT
    bCmdRun    : BOOL := FALSE; // 软启器运行端子输出（斜坡 / 旁路 / 运行相保持）[-] / the softstarter run terminal outlet
    bCmdBypass : BOOL := FALSE; // 旁路接触器线圈输出（仅投旁路与运行相）[-] / the bypass contactor coil outlet
END_VAR
VAR
    _ePhase    : E_DL_SsdPhase := E_DL_SsdPhase.eSsdIdle; // 内部相位，CASE 唯一写入目标 / the internal phase, the single CASE write target
    _uErrorId  : UDINT := 0;      // 内部故障码寄存（契约属性 uErrorId 数据源）/ the internal error register, the property data source
    _bFault    : BOOL := FALSE;   // 故障锁存位（契约属性 bFault 数据源之一）/ the fault latch bit
    _bCooling  : BOOL := FALSE;   // 冷却计时进行中 [-] / the cooling timing active
    _bInhibit  : BOOL := FALSE;   // 重启抑制激活寄存（契约属性 bRestartInhibit 数据源）/ the restart inhibit register
    _bPendStart: BOOL := FALSE;   // 方法启动请求（CmdStart 置位）/ the method start request
    _bPendReset: BOOL := FALSE;   // 方法复位请求（CmdReset 置位）/ the method reset request
    _bStopLatch: BOOL := FALSE;   // 停止锁存（引脚或方法置位，主体消化）/ the stop latch
    rtStart    : R_TRIG;          // 引脚启动指令沿，段 0 无条件刷新 / the pin start edge
    rtReset    : R_TRIG;          // 引脚复位沿，段 0 无条件刷新 / the pin reset edge
    tonRamp    : TON;             // 斜坡窗，段 0 无条件刷新 / the ramp window
    tonFb      : TON;             // 旁路反馈确认窗，段 0 无条件刷新 / the bypass feedback window
    tonStop    : TON;             // 停机分断确认窗，段 0 无条件刷新 / the stop confirm window
    tonInh     : TON;             // 重启抑制冷却窗，段 0 无条件刷新 / the restart inhibit cooling window
END_VAR

METHOD CmdStart : BOOL
VAR_INPUT
END_VAR
IF (_ePhase <> E_DL_SsdPhase.eSsdIdle) OR _bFault OR _bInhibit THEN // 非空闲 / 故障 / 抑制拒绝 / refused when not idle, faulty or inhibited
    CmdStart := FALSE; // 拒绝 / refused
ELSE // 受理 / accepted
    _bPendStart := TRUE; // 登记启动请求，主体状态机消化 / register the start request for the body
    CmdStart := TRUE; // 受理 / accepted
END_IF

(*------------------------------------------------------------------------------
 * 方法: CmdStop —— 无条件安全停止（双命令全断语义，主体在载能相消化）。
 *      Method CmdStop, the unconditional safe stop, consumed by the body in the powered phases.
 *------------------------------------------------------------------------------*)
    END_METHOD

METHOD CmdStop
VAR_INPUT
END_VAR
_bStopLatch := TRUE; // 登记停止锁存，主体状态机消化 / register the stop latch for the body

(*------------------------------------------------------------------------------
 * 方法: CmdReset —— 复位过载 / 故障，返回是否可复位。
 *      Method CmdReset, resets the overload or the fault, returns the resettable verdict.
 *------------------------------------------------------------------------------*)
    END_METHOD

METHOD CmdReset : BOOL
VAR_INPUT
END_VAR
IF _bFault OR (_ePhase = E_DL_SsdPhase.eSsdTrip) OR (_ePhase = E_DL_SsdPhase.eSsdFault) THEN // 存在锁存故障 / a latch exists
    _bPendReset := TRUE; // 登记复位请求，主体状态机消化 / register the reset request for the body
    CmdReset := TRUE; // 可复位 / resettable
ELSE // 无故障可复位 / nothing to reset
    CmdReset := FALSE; // 不可复位 / not resettable
END_IF

(*------------------------------------------------------------------------------
 * 属性: eState（GET）—— 当前状态（内部相位映射契约枚举 E_DL_MotorState）。
 *      Property eState, the internal phase mapped onto the contract enum.
 *------------------------------------------------------------------------------*)
    END_METHOD

// 段 0｜定时器与沿检测无条件周期刷新（禁入分支，FB50-1）/ segment 0, the unconditional refresh
rtStart(CLK := bCmdStart); // 启动沿 / the start edge
rtReset(CLK := bReset); // 复位沿 / the reset edge
tonRamp(IN := (_ePhase = E_DL_SsdPhase.eSsdRamp) AND (NOT _bFault), PT := tRampTime); // 斜坡窗，IN 串斜坡相闸 / the ramp window gated by the ramp phase
tonFb(IN := (_ePhase = E_DL_SsdPhase.eSsdByWait) AND (NOT _bFault), PT := tFbWindow); // 反馈窗，IN 串投旁路相闸 / the feedback window gated by the engage phase
tonStop(IN := (_ePhase = E_DL_SsdPhase.eSsdStop) AND (NOT _bFault), PT := tStopConfirm); // 停机窗，IN 串停机相闸 / the stop window gated by the stop phase
tonInh(IN := _bCooling, PT := tRestartInhibit); // 冷却窗自复位由到期分支消化 / the cooling window absorbed by the expiry branch
IF tonInh.Q THEN // 冷却到期 / the cooling expired
    _bCooling := FALSE; // 结束冷却计时 / stop the cooling timing
    _bInhibit := FALSE; // 解除重启抑制 / release the inhibit
ELSE // 冷却中 / while cooling
    _bInhibit := _bCooling; // 抑制寄存随冷却 / the inhibit follows the cooling
END_IF

// 段 1｜公约声明（本块为纯事件型状态机，无学习 / 积分 / 滤波状态，首扫跟踪
//       范式不适用，变量零值由编译器缺省保证，无内部初始化标志——与族内
//       FB_DL_DolMotor 公约 0.1 同口径）
// segment 1, the convention note, a pure event state machine with no learning or integral state

// 段 2｜复位沿作用域：清锁存 / 清码 / 迁空闲（三项逐项声明，R59 轻①：前置故障相位门——故障相位下复位只清锁存不迁相，
//       迁相交由 CASE 故障相复位分支消化，避免绕过 eSsdFault 分支的进冷却语义）/ segment 2, the reset edge scope
IF rtReset.Q THEN // 复位沿 / the reset edge
    IF _ePhase <> E_DL_SsdPhase.eSsdFault THEN // 故障相位门：非故障相才执行迁相 / the fault phase gate, migrate only outside the fault phase
        _bFault := FALSE; // 作用域一：清故障锁存 / scope one, clear the fault latch
        _uErrorId := 0; // 作用域二：清故障码 / scope two, clear the code
        _ePhase := E_DL_SsdPhase.eSsdIdle; // 作用域三：迁空闲相 / scope three, back to idle
    ELSE // 故障相位：仅清锁存与码，不迁相（迁相与进冷却由段 4 eSsdFault 分支消化）/ the fault phase, latch and code only
        _bFault := FALSE; // 清故障锁存 / clear the fault latch
        _uErrorId := 0; // 清故障码 / clear the code
    END_IF
END_IF

// 段 3｜过载全局监视（优先级最高，R190 独立成因独立码，边界三）/ segment 3, the global overload monitor
IF bOverload AND ((_ePhase = E_DL_SsdPhase.eSsdRamp) OR (_ePhase = E_DL_SsdPhase.eSsdByWait) OR (_ePhase = E_DL_SsdPhase.eSsdRun)) THEN // 载能相过载 / an overload in a powered phase
    _bFault  := TRUE; // 置故障锁存 / raise the fault latch
    _uErrorId := 16#0003_0215; // 0003_0215 过载锁存【故障级】/ the overload latch, fault grade
    _ePhase  := E_DL_SsdPhase.eSsdTrip; // 迁脱扣相（锁存与迁相同分支，FB50-1）/ migrate to the trip phase
END_IF

// 段 4｜相位机：ENUM + CASE，含 ELSE 非法相位兜底（R128）/ segment 4, the phase machine
CASE _ePhase OF

E_DL_SsdPhase.eSsdIdle: // 空闲相 / the idle phase
    IF _bStopLatch THEN // 停止锁存消化 / absorb the stop latch
        _bStopLatch := FALSE; // 锁存清零 / clear the latch
    END_IF
    IF _bPendStart OR rtStart.Q THEN // 启动请求 / a start request
        _bPendStart := FALSE; // 消费请求不自动重试 / consume the request, no retry
        IF bOverload THEN // 过载未复位静默拒绝（脱扣码已在过载相锁存，驻留不迁移）/ an overload present, silent refusal, dwell without migrate
        ELSIF NOT bPermitStart THEN // 联锁未满足静默拒绝（驻留不迁移，R59 轻②删自赋值死语句）/ the permit absent, silent refusal
        ELSIF _bInhibit THEN // 抑制期拒绝（信息级 0217，R190 独立成因，驻留不迁移）/ refused during the inhibit, info grade
            _uErrorId := 16#0003_0217; // 0003_0217 重启抑制期拒绝【信息级】/ the inhibit refusal, info grade
        ELSE // 受理启动 / accept the start
            _ePhase := E_DL_SsdPhase.eSsdRamp; // 迁斜坡相 / migrate to the ramp
        END_IF
    END_IF

E_DL_SsdPhase.eSsdRamp: // 斜坡相：运行端子得电旁路断开 / the ramp phase
    IF bFbBypass THEN // 旁路提前吸合矛盾（R190 独立成因）/ a premature bypass pick up contradiction
        _bFault  := TRUE; // 置故障锁存 / raise the fault latch
        _uErrorId := 16#0003_0214; // 0003_0214 斜坡期旁路提前吸合【故障级】/ the premature bypass, fault grade
        _ePhase  := E_DL_SsdPhase.eSsdFault; // 迁故障相 / migrate to the fault phase
    ELSIF bCmdStop OR _bStopLatch THEN // 停机中止 / a stop abort
        _bStopLatch := FALSE; // 消化停止锁存 / absorb the stop latch
        _ePhase := E_DL_SsdPhase.eSsdStop; // 迁停机相（启动中止无运行时长）/ migrate to the stop phase
    ELSIF tonRamp.Q THEN // 斜坡窗到 / the ramp done
        _ePhase := E_DL_SsdPhase.eSsdByWait; // 迁投旁路相 / migrate to the engage phase
    END_IF

E_DL_SsdPhase.eSsdByWait: // 投旁路相：等旁路反馈吸合确认 / the engage phase
    IF bFbBypass THEN // 反馈吸合确认 / the feedback confirmed
        _ePhase := E_DL_SsdPhase.eSsdRun; // 迁运行相 / migrate to the run phase
    ELSIF bCmdStop OR _bStopLatch THEN // 停机中止 / a stop abort
        _bStopLatch := FALSE; // 消化停止锁存 / absorb the stop latch
        _ePhase := E_DL_SsdPhase.eSsdStop; // 迁停机相 / migrate to the stop phase
    ELSIF tonFb.Q THEN // 反馈确认窗超时（启动超时保护）/ the feedback window timed out
        _bFault  := TRUE; // 置故障锁存 / raise the fault latch
        _uErrorId := 16#0003_0211; // 0003_0211 旁路反馈确认超时【故障级】/ the bypass feedback timeout, fault grade
        _ePhase  := E_DL_SsdPhase.eSsdFault; // 迁故障相 / migrate to the fault phase
    END_IF

E_DL_SsdPhase.eSsdRun: // 运行相：旁路反馈吸合确认带载 / the run phase
    IF NOT bFbBypass THEN // 运行中旁路反馈意外断开（R190 独立成因）/ the feedback dropped while running
        _bFault  := TRUE; // 置故障锁存 / raise the fault latch
        _uErrorId := 16#0003_0212; // 0003_0212 运行中旁路反馈断开【故障级】/ the feedback loss, fault grade
        _ePhase  := E_DL_SsdPhase.eSsdFault; // 迁故障相 / migrate to the fault phase
    ELSIF bCmdStop OR _bStopLatch THEN // 停机指令 / a stop command
        _bStopLatch := FALSE; // 消化停止锁存 / absorb the stop latch
        _ePhase := E_DL_SsdPhase.eSsdStop; // 迁停机相 / migrate to the stop phase
    END_IF

E_DL_SsdPhase.eSsdStop: // 停机过渡相：双命令全断等旁路分断确认（边界二）/ the stop transition phase
    IF NOT bFbBypass THEN // 旁路分断确认 / the drop out confirmed
        _bCooling := TRUE; // 启动重启抑制冷却 / start the cooling
        _ePhase := E_DL_SsdPhase.eSsdIdle; // 回空闲相 / back to idle
    ELSIF tonStop.Q THEN // 停机确认窗超时（触点粘连，R190 独立成因）/ the stop confirm timeout, a welded contact
        _bFault  := TRUE; // 置故障锁存 / raise the fault latch
        _uErrorId := 16#0003_0213; // 0003_0213 停机旁路未分断【故障级】/ the drop out timeout, fault grade
        _ePhase  := E_DL_SsdPhase.eSsdFault; // 迁故障相 / migrate to the fault phase
    END_IF

E_DL_SsdPhase.eSsdTrip: // 过载脱扣锁存相：仅复位且过载消失可清 / the trip latch phase
    IF (rtReset.Q OR _bPendReset) AND (NOT bOverload) THEN // 复位且过载消失 / a reset with the overload removed
        _bPendReset := FALSE; // 消费复位请求 / consume the reset request
        _bFault := FALSE; // 解除锁存（解除路径 = 复位沿，R188）/ release the latch
        _uErrorId := 0; // 清故障码 / clear the code
        _bCooling := TRUE; // 脱扣复位进冷却 / start the cooling
        _ePhase := E_DL_SsdPhase.eSsdIdle; // 回空闲相 / back to idle
    END_IF

E_DL_SsdPhase.eSsdFault: // 故障锁存相：仅复位可清 / the fault latch phase
    IF rtReset.Q OR _bPendReset THEN // 复位沿 / a reset edge
        _bPendReset := FALSE; // 消费复位请求 / consume the reset request
        _bFault := FALSE; // 解除锁存（解除路径 = 复位沿，R188）/ release the latch
        _uErrorId := 0; // 清故障码 / clear the code
        _bCooling := TRUE; // 故障复位进冷却 / start the cooling
        _ePhase := E_DL_SsdPhase.eSsdIdle; // 回空闲相 / back to idle
    END_IF

ELSE // 非法相位兜底（R128）/ the illegal phase fallback
    _bFault  := TRUE; // 置故障锁存 / raise the fault latch
    _uErrorId := 16#0003_0216; // 0003_0216 非法状态【故障级】/ the illegal state, fault grade
    _ePhase  := E_DL_SsdPhase.eSsdFault; // 迁故障相 / migrate to the fault phase
END_CASE

// 段 5｜统一出口：命令输出按相位单点映射（边界二安全侧全断）/ segment 5, the unified outlet
bCmdRun := (_ePhase = E_DL_SsdPhase.eSsdRamp) OR (_ePhase = E_DL_SsdPhase.eSsdByWait) OR (_ePhase = E_DL_SsdPhase.eSsdRun); // 运行端子仅载能相保持 / the run terminal held in the powered phases
bCmdBypass := (_ePhase = E_DL_SsdPhase.eSsdByWait) OR (_ePhase = E_DL_SsdPhase.eSsdRun); // 旁路线圈仅投旁路与运行相 / the bypass coil in the engage and run phases
IF _bFault OR (_ePhase = E_DL_SsdPhase.eSsdTrip) OR (_ePhase = E_DL_SsdPhase.eSsdFault) THEN // 故障相覆盖闸（R191 降级显式）/ the fault phase override
    bCmdRun := FALSE; // 运行端子安全侧断开 / the run terminal off on the safe side
    bCmdBypass := FALSE; // 旁路线圈安全侧断开 / the bypass coil off on the safe side
END_IF

(*------------------------------------------------------------------------------
 * 方法: CmdStart —— 启动指令（单发）。故障 / 脱扣 / 抑制 / 非空闲态返回 FALSE。
 *      Method CmdStart, a one shot start, FALSE when latched, tripped, inhibited or not idle.
 *------------------------------------------------------------------------------*)

PROPERTY eState : E_DL_MotorState
CASE _ePhase OF // 内部相位到契约枚举映射 / the internal phase to the contract enum mapping
E_DL_SsdPhase.eSsdIdle:   eState := E_DL_MotorState.eIdle;          // 空闲映射 / the idle mapping
E_DL_SsdPhase.eSsdRamp:   eState := E_DL_MotorState.eStarting;      // 斜坡归启动校验态 / the ramp mapped to starting
E_DL_SsdPhase.eSsdByWait: eState := E_DL_MotorState.eStarting;      // 投旁路归启动校验态 / the engage mapped to starting
E_DL_SsdPhase.eSsdRun:    eState := E_DL_MotorState.eRunning;       // 运行映射 / the run mapping
E_DL_SsdPhase.eSsdStop:   eState := E_DL_MotorState.eStopping;      // 停机映射 / the stop mapping
E_DL_SsdPhase.eSsdTrip:   eState := E_DL_MotorState.eTripOverload;  // 脱扣映射 / the trip mapping
E_DL_SsdPhase.eSsdFault:  eState := E_DL_MotorState.eFault;         // 故障映射 / the fault mapping
ELSE                      eState := E_DL_MotorState.eFault;         // 非法相位按故障态上报（R128）/ the illegal phase reported as the fault
END_CASE

(*------------------------------------------------------------------------------
 * 属性: bRunning（GET）—— 运行反馈（运行相且旁路反馈吸合确认）。
 *      Property bRunning, the run feedback, the run phase with the bypass confirmed.
 *------------------------------------------------------------------------------*)
PROPERTY bRunning : BOOL
bRunning := (_ePhase = E_DL_SsdPhase.eSsdRun) AND bFbBypass; // 显式确认式派生 / the explicit confirmed derived form

(*------------------------------------------------------------------------------
 * 属性: bFault（GET）—— 故障锁存指示（信息级 0217 不置本位，0.2 公约）。
 *      Property bFault, the fault latch indicator, the info code excluded.
 *------------------------------------------------------------------------------*)
PROPERTY bFault : BOOL
bFault := _bFault OR (_ePhase = E_DL_SsdPhase.eSsdTrip) OR (_ePhase = E_DL_SsdPhase.eSsdFault); // 显式排除信息级派生式 / the derived form excluding the info grade

(*------------------------------------------------------------------------------
 * 属性: uErrorId（GET）—— 末次故障码（0 = 无故障）。
 *      Property uErrorId, the last error code, zero when none.
 *------------------------------------------------------------------------------*)
PROPERTY uErrorId : UDINT
uErrorId := _uErrorId; // 返回内部故障码寄存 / return the internal error register

(*------------------------------------------------------------------------------
 * 属性: bRestartInhibit（GET）—— 重启抑制激活指示。
 *      Property bRestartInhibit, the restart inhibit active indicator.
 *------------------------------------------------------------------------------*)
PROPERTY bRestartInhibit : BOOL
bRestartInhibit := _bInhibit; // 返回抑制寄存 / return the inhibit register
END_FUNCTION_BLOCK

(* ---- FB_DL_SolenoidCoilHealth.st ---- *)
(*==============================================================================
 * 组件名称 (Component)  : FB_DL_SolenoidCoilHealth
 * 所属子库 (Sublibrary) : DL_Device
 * 当前版本 (Version)    : 1.0.0
 * 兼容性   (Platform)   : CODESYS 3.5+ / TwinCAT 3 / 汇川 InoProShop / 施耐德 Machine Expert
 *                         仅依赖 Standard.library（TON / R_TRIG / ABS），零厂商私有库
 * 功能描述 (Function)   : 电磁阀线圈电气健康诊断（吸合窗 / 保持段分域判据）：
 *                         ① 吸合窗：bEnergized 上升沿起 tWindow 内捕获峰值电流 fPickPeakA，
 *                            峰值 > fPickMaxA 判 eStuckPeak（衔铁卡阻 / 短路匝趋势）；
 *                         ② 保持段：窗后保持电流对学习基线 _fHoldBase 的偏差超 fHoldPct，
 *                            低偏判 eUnderCurrent（断匝趋势）、高偏判 eOverCurrent（短路匝
 *                            趋势）；基线自合格吸合（峰值入 [fPickMinA, fPickMaxA] 窗）递推
 *                            学习，n < 3 次合格吸合前**拒判**（不足拒判，防冷启动误报）。
 *                         ③ 电流 <= 0 且 bEnergized 持续 tWindow → eNoData（传感器断线，
 *                            不与欠流混码，R190 成因分码）。
 * 接口     (Interface)  : 输入 fCurrentA 线圈电流（A）、bEnergized 得电、tWindow 判据窗、
 *                         fPickMaxA/fPickMinA 吸合峰值窗（A）、fHoldPct 保持电流容差（%）、
 *                         bReset 复位；输出 eCoil 健康态、fPickPeakA 最近吸合峰值（A）、
 *                         bError 故障标志。
 * 边界     (Boundary)   : ① **属主边界（写死）：本件只做线圈电气健康诊断，不驱动线圈、
 *                         不判触点熔焊、不做阀通断动作**。
 *                         ② 非有限电流当拍剔除（不参与峰值与判据，R245）。
 *                         ③ 峰值窗 TON / 断线 TON 段 0 无条件刷新；IN 由状态表达式派生，
 *                         无外部沿清零。
 *                         ④ 组态闸：tWindow<=T#0S、fPickMaxA<=fPickMinA、fHoldPct<=0 →
 *                         锁存 bError 且 eCoil 冻结 eOk 侧不误报，解除沿 = bReset 上升沿。
 *                         ⑤ 基线递推：_fHoldBase += (窗末电流 - _fHoldBase)/_nPickOk
 *                         （均值增量式，_nPickOk 为 UDINT 合格吸合计数，饱和不回绕）。
 *                         ⑥ 每次得电下降沿回 eOff 并清吸合窗标志；诊断态在失电后不保持
 *                         （健康态按周期重判）。
 *                         ⑦ 零全局耦合（无 GVL / 无 VAR_EXTERNAL / 无物理地址）。
 * 分工声明 (Scope)      : 与 `FB_DL_ContactorWeldDetect` 分工：线圈电气健康（本件）≠ 触点
 *                         熔焊（那件）；与 `FB_DL_SingleSolenoidCyl` 分工：诊断 ≠ 通断驱动。
 * 来源标签 (Source Tag) : T2-6 ◐（Rockwell AOI 设备诊断粒度只借"吸合窗/保持段分域"分类
 *                         事实，判据与基线学习为本件自研实现）
 * 码表     (Codes)      : 本件不占用任何全局数字码位。出口为 ENUM 健康态 + LREAL 峰值 +
 *                         BOOL；数字码位待主控收口阶段统一派号。
 * 红线自检 (Redline)    : R1 ✓ 零 GVL/VAR_EXTERNAL ｜ R2 ✓ 零 %I/%Q/%M ｜ R3 ✓ 纯 IEC 61131-3
 *                         R4 ✓ 除零前置（均值分母计数闸）+ 非有限剔除 + 组态闸 ｜ R5 ✓ 声明逐行同行双语注释
 *                         R6 ✓ ENUM 健康态 CASE 化判序 ｜ R7 ✓ 两 TON/两 R_TRIG 段 0 无条件刷新
 * 修订历史 (Revision)   : 2026-11-20  v1.0.0  R48 首版（批次 2 · 序号 10）
 *                         验收向量：峰值超上限 → eStuckPeak；保持欠偏 → eUnderCurrent；
 *                         电流恒 0 得电 → eNoData；n<3 合格吸合 → 拒判 eOk。
 *==============================================================================*)

TYPE E_DL_SchHealth :
(
    eOk           := 0,    // 健康（含拒判期）/ Healthy, including not-yet-judged period
    eUnderCurrent := 10,   // 保持欠流（断匝趋势）/ Hold under-current, turn-short-open trend
    eOverCurrent  := 20,   // 保持过流（短路匝趋势）/ Hold over-current, turn-short trend
    eStuckPeak    := 30,   // 吸合峰值超上限（衔铁卡阻）/ Pickup peak above ceiling, armature stuck
    eNoData       := 40,   // 传感器断线（得电而电流恒零）/ No data, sensor dead while energized
    eOff          := 50    // 线圈失电（判据冻结）/ Coil de-energized, judges frozen
);
END_TYPE

FUNCTION_BLOCK FB_DL_SolenoidCoilHealth
VAR_INPUT
    fCurrentA : LREAL := 0.0;    // 线圈电流实测 [A] / Coil current measurement [A]
    bEnergized: BOOL := FALSE;   // 线圈得电命令反馈 [-] / Coil energized state
    tWindow   : TIME := T#500MS; // 吸合判据窗（峰值捕获与断线判据共用窗长），域 > T#0S [ms] / Pickup judge window [ms]
    fPickMaxA : LREAL := 2.0;    // 吸合峰值窗上限，域 > fPickMinA [A] / Pickup peak window ceiling [A]
    fPickMinA : LREAL := 1.0;    // 吸合峰值窗下限，域 >= 0 [A] / Pickup peak window floor [A]
    fHoldPct  : LREAL := 20.0;   // 保持电流容差（对基线百分比），域 > 0 [%] / Hold current tolerance vs baseline [%]
    bReset    : BOOL := FALSE;   // 复位，上升沿清组态故障锁存 [-] / Reset, rising edge clears config latch
END_VAR
VAR_OUTPUT
    eCoil      : E_DL_SchHealth;  // 线圈健康态出口 [-] / Coil health outlet
    fPickPeakA : LREAL;            // 最近一次吸合峰值电流（失电保持供诊断） [A] / Last captured pickup peak [A]
    bError     : BOOL;            // 故障标志（组态非法 ∨ 健康态非 eOk/eOff） [-] / Error flag
END_VAR
VAR
    _eCoil    : E_DL_SchHealth := E_DL_SchHealth.eOff;   // 内部健康态 / Internal health state
    _bPickWin : BOOL;               // 吸合窗开启标志（上升沿置位、窗到清除） / Pickup window open flag
    _fPeak    : LREAL := 0.0;       // 当次吸合峰值跟踪 [A] / Current pickup peak tracker
    _fHoldBase: LREAL := 0.0;       // 保持电流学习基线（递推均值） [A] / Learned hold-current baseline
    _nPickOk  : UDINT := 0;         // 合格吸合计数（基线判据门槛 n>=3，诊断用） [次] / Qualified pickup count
    _nDiv     : LREAL := 0.0;       // 均值递推实数除数（随合格吸合递增，判零前置） / Mean recursion real divisor
    _fDevLim  : LREAL;              // 保持段容差绝对限（基线×fHoldPct） [A] / Hold tolerance absolute limit
    _bErrLatch: BOOL;               // 组态故障锁存位（解除沿 = bReset 上升沿） / Latched config fault, cleared by reset edge
    tonPickWin: TON;                // 吸合峰值窗定时器，段 0 无条件调用 / Pickup window timer
    tonNoData : TON;                // 断线判据定时器，段 0 无条件调用 / No-data timer
    rtEn      : R_TRIG;             // 得电上升沿实例，段 0 无条件调用 / Energize rising edge instance
    rtDis     : R_TRIG;             // 失电下降沿实例（F_TRIG 语义由 R_TRIG 反相实现），段 0 无条件调用 / De-energize falling edge instance
    rtReset   : R_TRIG;             // 复位沿实例，段 0 无条件调用 / Reset edge instance
    _bNonFin  : BOOL;               // 电流非有限当拍量 [-] / Non-finite current this scan
END_VAR
VAR CONSTANT
    DL_SCH_UDMAX   : UDINT := 4294967295;   // UDINT 上限（合格吸合计数饱和点） [次] / UDINT ceiling for count saturation
    DL_SCH_NMIN    : UDINT := 3;            // 基线生效最小合格吸合次数 [次] / Minimum qualified pickups for baseline
    DL_SCH_ZEROTH  : LREAL := 0.0;          // 电流判零基准（断线判据） [A] / Current zero base for no-data test
    DL_SCH_EPS     : LREAL := 0.0;          // 非有限差值判零基准 [-] / Non-finite difference zero base
    DL_SCH_PCT     : LREAL := 100.0;        // 百分比换算基 [无量纲] / Percent conversion base
END_VAR

(* —— 段 0：非有限判 + 组态闸 + 两 TON 三沿无条件周期刷新 —— *)
_bNonFin := (fCurrentA <> fCurrentA) OR ((fCurrentA - fCurrentA) <> DL_SCH_EPS);   // 电流非有限（R245） / Non-finite current
IF (tWindow <= T#0S) OR (fPickMaxA <= fPickMinA) OR (fPickMinA < DL_SCH_ZEROTH) OR (fHoldPct <= 0.0) THEN
    _bErrLatch := TRUE;                                     // 组态域闸：锁存（R188 解除沿 = bReset 上升沿） / Config gate: latch
END_IF
rtEn(CLK := bEnergized);                                    // 得电沿，每拍必调 / Energize edge, every scan
rtDis(CLK := NOT bEnergized);                               // 失电沿（反相实现下降沿），每拍必调 / De-energize edge, every scan
rtReset(CLK := bReset);                                     // 复位沿，每拍必调 / Reset edge, every scan
tonPickWin(IN := _bPickWin, PT := tWindow);                 // 吸合峰值窗（IN 状态派生，无外部清零） / Pickup window timer
tonNoData(IN := bEnergized AND (fCurrentA <= DL_SCH_ZEROTH) AND (NOT _bNonFin), PT := tWindow);   // 断线判据窗 / No-data judge window

(* —— 段 1：复位沿 / 失电沿（窗态与判据态清出） —— *)
IF rtReset.Q THEN
    _bErrLatch := FALSE;                                    // 清组态故障锁存 / Clear config latch
END_IF
IF rtDis.Q THEN
    _bPickWin := FALSE;                                     // 失电关吸合窗 / Close pickup window on de-energize
    _eCoil := E_DL_SchHealth.eOff;                          // 失电判据冻结回 eOff / Freeze to eOff
END_IF

(* —— 段 2：吸合窗开启与峰值捕获 —— *)
IF rtEn.Q THEN
    _bPickWin := TRUE;                                      // 得电沿开启吸合窗 / Open pickup window on energize edge
    _fPeak := 0.0;                                          // 峰值跟踪清零重捕 / Reset peak tracker
END_IF
IF _bPickWin AND (NOT _bNonFin) THEN
    IF fCurrentA > _fPeak THEN
        _fPeak := fCurrentA;                                // 峰值捕获（正电流单调上取） / Capture peak
    END_IF
END_IF

(* —— 段 3：窗到裁决（判吸合窗 → 基线学习） —— *)
IF tonPickWin.Q THEN
    _bPickWin := FALSE;                                     // 窗到关闭（下一拍 IN 派生自复位） / Close window at Q
    IF _fPeak > fPickMaxA THEN
        _eCoil := E_DL_SchHealth.eStuckPeak;                // 峰值超上限：判卡阻（R190 独立成因） / Peak above ceiling: stuck
    ELSIF _fPeak >= fPickMinA THEN
        IF _nPickOk < DL_SCH_UDMAX THEN
            _nPickOk := _nPickOk + 1;                       // 合格吸合计数（饱和不回绕） / Count qualified pickup, saturating
        END_IF
        _nDiv := _nDiv + 1.0;                               // 实数除数同步递增（避免 UDINT 转型溢出） / Real divisor increments in step
        IF (NOT _bNonFin) AND (_nDiv >= 1.0) THEN
            _fHoldBase := _fHoldBase + (fCurrentA - _fHoldBase) / _nDiv;   // 基线增量均值学习（除数恒 >=1） / Incremental mean baseline learning
        END_IF
        (* 合格吸合当拍不直接判健康，进入保持段分域判据（段 4） *)
        _eCoil := E_DL_SchHealth.eOk;                       // 吸合窗内默认健康（保持段再判） / Default healthy in window
    ELSE
        _eCoil := E_DL_SchHealth.eOk;                       // 峰值偏弱不判卡阻不学基线（保持段判欠流） / Weak peak: left to hold judge
    END_IF
END_IF

(* —— 段 4：保持段判据（窗后得电期；n<3 拒判） —— *)
IF bEnergized AND (NOT _bPickWin) AND (NOT _bErrLatch) THEN
    IF tonNoData.Q THEN
        _eCoil := E_DL_SchHealth.eNoData;                   // 电流恒零：传感器断线（不与欠流混码，R190） / Constant zero current: no data
    ELSIF _nPickOk >= DL_SCH_NMIN THEN
        _fDevLim := _fHoldBase * fHoldPct / DL_SCH_PCT;     // 保持容差绝对限 [A] / Hold tolerance absolute limit
        IF (fCurrentA < _fHoldBase - _fDevLim) AND (NOT _bNonFin) THEN
            _eCoil := E_DL_SchHealth.eUnderCurrent;         // 欠偏：断匝趋势 / Under deviation: open-turn trend
        ELSIF (fCurrentA > _fHoldBase + _fDevLim) AND (NOT _bNonFin) THEN
            _eCoil := E_DL_SchHealth.eOverCurrent;          // 过偏：短路匝趋势 / Over deviation: short-turn trend
        ELSE
            _eCoil := E_DL_SchHealth.eOk;                   // 带内健康 / In-band healthy
        END_IF
    ELSE
        _eCoil := E_DL_SchHealth.eOk;                       // 合格吸合不足 3 次：拒判（防冷启动误报） / Fewer than three pickups: not judged
    END_IF
END_IF

(* —— 段 5：出口单点映射（名实双出口同源，R191） —— *)
eCoil := _eCoil;                                            // 健康态出口 / Health outlet
fPickPeakA := _fPeak;                                       // 最近吸合峰值出口（失电保持供诊断） / Last peak outlet, kept on de-energize
bError := _bErrLatch
       OR (_eCoil = E_DL_SchHealth.eNoData)
       OR (_eCoil = E_DL_SchHealth.eStuckPeak)
       OR (_eCoil = E_DL_SchHealth.eOverCurrent)
       OR (_eCoil = E_DL_SchHealth.eUnderCurrent);          // 故障标志 = 组态非法 ∨ 任一非健康态（与 eCoil 同源配对） / Error = cfg fault or any unhealthy state

END_FUNCTION_BLOCK

(* ---- FB_DL_SprayNozzleBank.st ---- *)
(*
  ==================================================================
  组件名 Component  : FB_DL_SprayNozzleBank
  分类   Category   : DL_Device
  复杂度 Complexity  : 中
  版本   Version    : 1.0.0
  功能   Purpose    : 多喷嘴组排布时序（8 组上限）。分段分组吹扫/喷涂：组
                      计时 tGroup 到迁下一组，组间搭接窗 tOverlap 内前组维
                      持得电；喷堵压力反馈诊断：组活动期压力持续超阈值计满
                      tClogMon 判喷堵，累计 nClogCnt 达限锁存报警。LBP 命令
                      → 监视 → 判定骨架。
  来源   Source     : T2-2-lbp（命令→监视→判定骨架）
  溯源   Origin     : IEC 61131-3 标准语义的道莅防御性实现；喷嘴分组时序与
                      压差诊断为行业公知工程语义，clean-room 自研实现，未复
                      制 LBP 或任何厂商私有库源码。
  平台   Platform   : 纯 IEC 61131-3（Standard.library: TON / R_TRIG，无私有库）
  分工声明 Split     : 与 FB_DL_DustCollectorPulse 分工——后者做除尘脉冲轮
                      巡反吹，本件做喷嘴组搭接排布时序。
  作者   Author     : 道莅代码库 · PLC 编程专家（R59）
  ------------------------------------------------------------------
  边界 Boundary     :
                      一 安全语义：停机 / 故障 / 喷堵报警 / 非有限压力时全组
                         输出统一出口强制 FALSE（安全侧单点映射，R191）；
                      二 组态域闸：nGroups ∈ [1..8]，越域锁存 bError（解除
                         = bReset 沿，R188）；
                      三 搭接窗 tOverlap < tGroup 由调用方保证，本件不二次
                         钳制；组计时窗到期即迁（窗口末退出迁移，纪律④）；
                      四 喷堵诊断：非有限压力置 bBad 挂起监视（不误报不吞），
                         组活动期 tonClog 计满判堵一次计数（自复位窗，R188）；
                      五 定时器与沿检测全部段 0 无条件周期刷新（R7）；
                      六 无全局变量、无外部变量声明、无物理地址寻址。
  修订记录 Revision  :
    2026-11-21  v1.0.0  R59 首版（批 2 · 序号 9）
  ==================================================================
*)

TYPE E_DL_SnbPhase :
(
    eSnbIdle := 0,  // 空闲：消化停止与复位 / idle, absorbing the stop and reset
    eSnbRun  := 10, // 分组排布运行：组计时推进 / the group sequencing run
    eSnbDone := 20, // 全组完成驻留：等新启动沿 / the all groups done dwell
    eSnbFault := 90 // 故障锁存：仅复位可清 / the latched fault
);
END_TYPE

FUNCTION_BLOCK FB_DL_SprayNozzleBank
VAR_INPUT
    bStart     : BOOL := FALSE; // 启动指令，上升沿生效 [-] / the start command, rising edge effective
    bStop      : BOOL := FALSE; // 停止指令，电平生效 [-] / the stop command, level effective
    nGroups    : INT  := 8;     // 组数组态 [组]，域 1..8 / the group count config, one through eight
    tGroup     : TIME := T#2S;  // 单组作用时长 [毫秒] / the per group duration [millisecond]
    tOverlap   : TIME := T#200MS; // 组间搭接窗 [毫秒] / the group overlap window [millisecond]
    fPress     : LREAL := 0.0;  // 喷嘴压力反馈 [千帕] / the nozzle pressure feedback [kilopascal]
    fPressClog : LREAL := 300.0; // 喷堵压力阈值 [千帕] / the clog pressure threshold [kilopascal]
    tClogMon   : TIME := T#1S;  // 喷堵判满窗（压力超阈值持续时长）[毫秒] / the clog verdict window [millisecond]
    nClogMax   : UDINT := 5;    // 喷堵计数报警限 [次] / the clog count alarm bound
    bReset     : BOOL := FALSE; // 报警与故障复位，上升沿生效 [-] / the alarm and fault reset, rising edge
END_VAR
VAR_OUTPUT
    aGrp     : ARRAY[0..7] OF BOOL; // 组输出组（仅前 nGroups 组参与排布）[-] / the group outlets
    nGrpIdx  : INT  := -1;  // 当前活动组索引，-1 = 无 [组] / the active group index, minus one when none
    bRunning : BOOL := FALSE; // 排布运行指示 [-] / the sequencing running indicator
    bDone    : BOOL := FALSE; // 全组完成单脉冲（单拍）[-] / the all done one shot pulse, single scan
    bClogAlm : BOOL := FALSE; // 喷堵报警锁存（解除 = bReset 沿）[-] / the clog alarm latch, released by the reset edge
    nClogCnt : UDINT := 0;    // 喷堵判定累计 [次] / the clog verdict count
    bBad     : BOOL := FALSE; // 非有限压力实时标志 [-] / the non finite pressure flag
    bError   : BOOL := FALSE; // 组态域闸故障锁存 [-] / the config gate fault latch
END_VAR
VAR CONSTANT
    DL_SNB_GRPMAX  : INT  := 8;          // 组容量上界 [组] / the group capacity bound
    DL_SNB_CNTMAX  : UDINT := 4294967294; // 计数防回绕上界 [次] / the counter anti wrap clamp bound
END_VAR
VAR
    _ePhase  : E_DL_SnbPhase := E_DL_SnbPhase.eSnbIdle; // 内部相位，CASE 唯一写入目标 / the internal phase, the single CASE write target
    _nGrp    : INT := 0;   // 组推进寄存 [组] / the group advance register
    _nI      : DINT;       // 组遍历索引（清零与出口重映射环）/ the group loop index
    _bOvlRun : BOOL := FALSE; // 搭接窗进行寄存（前组维持得电源）/ the overlap window register
    _bAdv    : BOOL := FALSE; // 组推进屏蔽寄存（组计时器重启一拍用）/ the advance mask register, the timer restart mask
    _bInit   : BOOL := FALSE; // 首拍初始化标志（R310，真实使用：首拍清组输出）/ the first scan flag, real use
    _bFinP   : BOOL;        // 压力有限工作量 [-] / the pressure finiteness work flag
    rtStart  : R_TRIG;      // 启动沿，段 0 无条件刷新 / the start edge
    rtReset  : R_TRIG;      // 复位沿，段 0 无条件刷新 / the reset edge
    tonGrp   : TON;         // 组计时窗，段 0 无条件刷新 / the group window
    tonOvl   : TON;         // 搭接窗（自复位一次性），段 0 无条件刷新 / the overlap one shot window
    tonClog  : TON;         // 喷堵判满窗（自复位），段 0 无条件刷新 / the clog verdict self reset window
END_VAR

// 段 0｜定时器与沿检测无条件周期刷新（禁入分支，R7）/ segment 0, the unconditional refresh
rtStart(CLK := bStart); // 启动沿 / the start edge
rtReset(CLK := bReset); // 复位沿 / the reset edge
tonGrp(IN := (_ePhase = E_DL_SnbPhase.eSnbRun) AND (NOT _bAdv), PT := tGroup); // 组计时窗，推进屏蔽一拍 / the group window, masked one scan per advance
tonOvl(IN := _bOvlRun, PT := tOverlap); // 搭接窗 / the overlap window
tonClog(IN := (_ePhase = E_DL_SnbPhase.eSnbRun) AND (NOT tonClog.Q) AND _bFinP AND (fPress > fPressClog), PT := tClogMon); // 自复位喷堵窗（R188）/ the self reset clog window

// 段 1｜首拍初始化（R310 真实使用路径）：组输出显式清零 / segment 1, the first scan init
IF NOT _bInit THEN // 首拍一拍 / the first scan
    _bInit := TRUE; // 置首拍标志 / raise the flag
    FOR _nI := 0 TO DL_SNB_GRPMAX - 1 DO // 全组清零 / clear all the groups
        aGrp[_nI] := FALSE; // 组输出清零 / clear the group outlet
    END_FOR
END_IF

// 段 2｜组态域闸与复位（边界二，解除路径 = bReset 沿，R188）/ segment 2, the config gate and the reset
IF (nGroups < 1) OR (nGroups > DL_SNB_GRPMAX) THEN // 组数越域 / the group count out of domain
    bError := TRUE; // 置域闸故障锁存 / raise the config latch
END_IF
IF rtReset.Q THEN // 复位沿 / the reset edge
    bError := FALSE; // 清域闸锁存 / clear the config latch
    bClogAlm := FALSE; // 清喷堵报警（解除路径声明）/ clear the clog alarm
    nClogCnt := 0; // 清喷堵计数 / clear the clog count
END_IF

// 段 3｜压力有限性与喷堵计数（非有限挂起监视不误报，边界四）/ segment 3, the pressure finiteness and the clog count
_bFinP := (fPress = fPress) AND ((fPress - fPress) = (fPress - fPress)); // 压力有限双判据（R79）/ the finiteness dual verdicts
bBad := NOT _bFinP; // 拒收实时标志与工作量同源（R191 名实双出口）/ the rejection flag shares the work flag
IF tonClog.Q THEN // 喷堵判满窗到期 / the clog window expired
    IF nClogCnt < DL_SNB_CNTMAX THEN // 计数防回绕 / the wrap guard
        nClogCnt := nClogCnt + 1; // 计一次 / count one
    END_IF
    IF nClogCnt >= nClogMax THEN // 达报警限 / at the alarm bound
        bClogAlm := TRUE; // 置喷堵报警锁存 / raise the clog alarm latch
    END_IF
END_IF

// 段 4｜单拍脉冲预清零（本库纪律③）/ segment 4, the per scan pulse preset
bDone := FALSE; // 完成脉冲预清零 / preset the done pulse false

// 段 5｜相位机：ENUM + CASE，含 ELSE 非法相位兜底（R6 / R128）/ segment 5, the phase machine
CASE _ePhase OF

E_DL_SnbPhase.eSnbIdle: // 空闲相 / the idle phase
    IF bStop THEN _nGrp := 0; END_IF // 停止消化（安全侧已在出口） / absorb the stop
    IF rtStart.Q AND (NOT bError) AND (NOT bClogAlm) THEN // 受理启动（组态合法且无报警）/ accept the start
        _nGrp := 0; // 组归零 / reset the group
        _ePhase := E_DL_SnbPhase.eSnbRun; // 运行相 / to the run phase
    END_IF

E_DL_SnbPhase.eSnbRun: // 排布运行相 / the run phase
    IF bStop OR bError OR bClogAlm THEN // 停止 / 组态故障 / 报警中止 / a stop, config fault or alarm abort
        _ePhase := E_DL_SnbPhase.eSnbIdle; // 回空闲 / back to idle
        _bOvlRun := FALSE; // 搭接窗取消 / cancel the overlap
    ELSE // 正常推进 / the normal advance
        IF tonGrp.Q THEN // 组计时窗到期（窗口末退出迁移，边界三）/ the group window expired
            _bAdv := TRUE; // 推进屏蔽一拍（组计时器下拍重启）/ raise the advance mask
            IF _nGrp > 0 THEN // 非首组：开启搭接窗维持前组 / a later group, open the overlap for the former
                _bOvlRun := TRUE; // 搭接窗启动 / start the overlap
            END_IF
            _nGrp := _nGrp + 1; // 组推进 / advance the group
            IF _nGrp >= nGroups THEN // 全组完成 / all the groups done
                _nGrp := 0; // 组归零 / reset the group
                _ePhase := E_DL_SnbPhase.eSnbDone; // 完成驻留相 / to the done dwell
                bDone := TRUE; // 置完成单脉冲 / raise the done pulse
            END_IF
        END_IF
    END_IF

E_DL_SnbPhase.eSnbDone: // 完成驻留相 / the done dwell phase
    IF bStop THEN // 停止消化 / absorb the stop
        _ePhase := E_DL_SnbPhase.eSnbIdle; // 回空闲 / back to idle
    END_IF

E_DL_SnbPhase.eSnbFault: // 故障锁存相（本件当前无迁入源，保留兜底对称位）/ the fault latch phase, reserved symmetric
    IF rtReset.Q THEN // 复位沿 / the reset edge
        _ePhase := E_DL_SnbPhase.eSnbIdle; // 回空闲 / back to idle
    END_IF

ELSE // 非法相位兜底（R128）/ the illegal phase fallback
    _ePhase := E_DL_SnbPhase.eSnbIdle; // 回空闲安全相 / back to the safe idle
END_CASE

// 段 6｜搭接窗消化与推进屏蔽清除（每拍后段执行）/ segment 6, the overlap consume and the mask clear
IF tonOvl.Q THEN // 搭接窗到期（窗口末退出）/ the overlap expired
    _bOvlRun := FALSE; // 前组断电 / drop the former group
END_IF
_bAdv := FALSE; // 推进屏蔽每拍清（组计时器重启机制）/ clear the advance mask every scan

// 段 7｜统一出口：组输出单点安全映射（边界一）/ segment 7, the unified outlet
FOR _nI := 0 TO DL_SNB_GRPMAX - 1 DO // 全组重映射 / remap all the groups
    aGrp[_nI] := FALSE; // 先全断（安全侧基线）/ all off first, the safe baseline
END_FOR
IF (_ePhase = E_DL_SnbPhase.eSnbRun) AND (NOT bError) AND (NOT bClogAlm) AND (NOT bStop) THEN // 排布有效窗口 / the valid sequencing window
    IF (_nGrp >= 0) AND (_nGrp < nGroups) THEN // 组界闸（防越界写）/ the group bound gate
        aGrp[_nGrp] := TRUE; // 当前组得电 / the current group on
    END_IF
    IF _bOvlRun AND (_nGrp > 0) AND (_nGrp - 1 < nGroups) THEN // 搭接窗内前组维持（组界闸）/ the former group held in the overlap
        aGrp[_nGrp - 1] := TRUE; // 前组得电 / the former group on
    END_IF
END_IF
nGrpIdx := _nGrp; // 活动组出口 / the active group outlet
bRunning := (_ePhase = E_DL_SnbPhase.eSnbRun); // 运行指示（R191 名实双出口）/ the running indicator
END_FUNCTION_BLOCK

(* ---- FB_DL_SsrHeaterDrive.st ---- *)
(*
    FB_DL_SsrHeaterDrive —— 固态继电器加热驱动
    ------------------------------------------------------------------
    分类      : DL_Device / Drive
    前缀      : FB_DL_
    版本      : 1.0.0
    溯源      : T2-2 LBP（只借「驱动块参数化 = 给定 + 周期 + 反馈诊断」的组内组织方式）；
                PWM 相位逻辑、断线判据、码位与分级 100% 自有；clean-room 重写，
                未复制任何闭源厂商源码，参考实现仅限 MIT/Apache 许可
    平台      : 纯 IEC 61131-3，CODESYS V3.5+ / TwinCAT 3 / InoProShop 通用
    作者      : 道莅代码库 · PLC编程专家（R18）
    ------------------------------------------------------------------
    功能说明  : 把连续功率需求 0~100 % 变成周期 PWM 的通断指令，并在「占空比足量却测
                不到加热电流」时判 SSR 开路 / 加热丝断线——这是本件的核心诊断，现场
                SSR 击穿或开路只表现为「温度不升」，没有电流检测永远查不出来；
                过零同步不做电网采样（零厂商依赖），改为「周期起点对齐 + 上层可注入
                同步脉冲」的声明式设计；
                三道闸：周期参数闸（周期非法时宁可断热，绝不满功率长通）→ 占空钳位闸
                → 零占空不启电流监视闸（零占空本来就没电流，否则误报）；
                时间比较全程用 TIME 原值，不转 REAL，避免毫秒精度损失。
    错误码    : 16#0003_0168 功率需求超域已钳位 / 占空低于导通阈值强制断——信息级，不置故障
                16#0003_0169 预留禁用（信息级，不得挪用）
                16#0003_032D PWM 周期参数非法，输出强制断开——故障级
                16#0003_032E 加热回路开路（占空足量但无电流超确认窗），锁存——故障级
                16#0003_032F 预留禁用（故障级，不得挪用）
    码位总账  : 16#0003_0168 用 / 16#0003_0169 预留 ｜ 16#0003_032D 用 / 16#0003_032E 用 / 16#0003_032F 预留
    状态机    : 无 CASE，周期相位由 TON 承载；bLoadLatch 为锁存位，非法状态不可能出现
    采样约定  : fbCycle / fbNoCurrent 与两个 R_TRIG 在本体首部无条件调用；tCycleTime
                必须与被控对象热惯性匹配，周期过短会让 SSR 频繁通断、寿命下降。
    修订记录  : 2026-11-16 v1.0.0 首次入库（R18）
*)
FUNCTION_BLOCK FB_DL_SsrHeaterDrive
VAR_INPUT
    bEnable            : BOOL;                 // 使能，FALSE 强制断输出（安全侧）/ enable, FALSE forces the output off, safe side
    bReset             : BOOL;                 // 上升沿清断线锁存 / rising edge clears the open circuit latch
    fPowerDemand       : REAL := 0.0;          // 功率需求 [%]，范围 0.0~100.0，超域钳位 / power demand [%], range 0.0~100.0, clamped outside
    tCycleTime         : TIME := T#1S;         // PWM 周期 [ms]，范围 500~10000 / PWM period [ms], range 500~10000
    bCurrentFeedback   : BOOL := FALSE;        // 加热电流检测输入，TRUE = 有电流 / heating current detection input, TRUE = current flows
    fMinDutyForCurrent : REAL := 10.0;         // 判定应有电流的最小占空 [%]，范围 1.0~50.0 / minimum duty that should produce current [%], range 1.0~50.0
    tCurrentWindow     : TIME := T#3S;         // 电流缺失确认窗 [ms]，范围 100~30000 / current absence confirmation window [ms], range 100~30000
    bSyncPulse         : BOOL := FALSE;        // 可选过零 / 同步脉冲，上升沿对齐周期起点 / optional zero crossing pulse, its rising edge aligns the cycle start
END_VAR
VAR_OUTPUT
    bOut         : BOOL;                       // SSR 驱动输出，TRUE = 导通 / SSR drive output, TRUE = conducting
    fDutyApplied : REAL;                       // 实际生效占空，钳位后 [%] / effective duty after clamping [%]
    tOnTime      : TIME;                       // 本周期已导通时长 [ms] / conducted time inside the current cycle [ms]
    bLoadOpen    : BOOL;                       // 加热回路开路，锁存，需复位 / heating circuit open, latched until reset
    eErr         : UDINT;                      // 错误码，0=正常 / error id, 0=ok
    bError       : BOOL;                       // 故障标志，eErr 为故障级时 TRUE / error flag, TRUE on fault-level eErr
END_VAR
VAR
    fbTrigReset  : R_TRIG;                     // 复位沿检测实例，本体首部无条件刷新 / reset edge instance, refreshed unconditionally
    fbTrigSync   : R_TRIG;                     // 同步脉冲沿检测实例，本体首部无条件刷新 / sync pulse edge instance, refreshed unconditionally
    fbCycle      : TON;                        // 周期相位定时器，自复位产生锯齿相位 / cycle phase timer, self-resetting to form a sawtooth phase
    fbNoCurrent  : TON;                        // 电流缺失确认定时器，本体首部无条件刷新 / current absence confirmation timer, refreshed unconditionally
    bCycleHold   : BOOL;                       // 周期相位保持位，IN 取反本定时器输出实现自复位 / phase hold bit, the inverted timer output self-resets it
    bForceRestart: BOOL;                       // 同步强制重启标志，单拍 / forced restart flag from the sync pulse, single cycle
    fDutyEff     : REAL;                       // 生效占空，钳位后 [%] / effective duty after clamping [%]
    fMinDutyEff  : REAL;                       // 生效电流判定最小占空，钳位后 [%] / effective minimum duty for the current check [%]
    tWindowEff   : TIME;                       // 生效电流确认窗，钳位后 [ms] / effective current confirmation window [ms]
    fCycleMs     : REAL;                       // 周期毫秒值，仅用于换算导通目标 [ms] / cycle in milliseconds, used for the on target only [ms]
    tOnTarget    : TIME;                       // 本周期应导通时长 [ms] / target conducted time inside the cycle [ms]
    fOnMs        : REAL;                       // 应导通时长的毫秒中间量 [ms] / target conducted time in milliseconds [ms]
    bLoadLatch   : BOOL;                       // 断线锁存位，仅复位清除 / open circuit latch, cleared by reset only
END_VAR
VAR CONSTANT
    DL_SSR_CYCLE_MIN  : TIME := T#500MS;       // PWM 周期下限 [ms] / PWM period lower bound [ms]
    DL_SSR_CYCLE_MAX  : TIME := T#10S;         // PWM 周期上限 [ms] / PWM period upper bound [ms]
    DL_SSR_WIN_MIN    : TIME := T#100MS;       // 电流确认窗下限 [ms] / current window lower bound [ms]
    DL_SSR_WIN_MAX    : TIME := T#30S;         // 电流确认窗上限 [ms] / current window upper bound [ms]
    DL_SSR_DUTY_MAX   : REAL := 100.0;         // 占空上限 [%] / duty upper bound [%]
    DL_SSR_DUTY_MIN   : REAL := 0.0;           // 占空下限 [%] / duty lower bound [%]
    DL_SSR_ON_EPS     : REAL := 0.5;           // 占空小于此视为全断 [%] / duties below this count as fully off [%]
    DL_SSR_MIND_MIN   : REAL := 1.0;           // 最小电流占空下限 [%] / minimum current duty lower bound [%]
    DL_SSR_MIND_MAX   : REAL := 50.0;          // 最小电流占空上限 [%] / minimum current duty upper bound [%]
    DL_SSR_PCT_SCALE  : REAL := 100.0;         // 百分比换算除数，恒非零 [%] / percentage scaling divisor, never zero [%]
    DL_FLOAT_EPS      : REAL := 1.0E-6;        // 浮点判等容差 [%] / float equality tolerance [%]
    DL_SSR_ZERO_REAL  : REAL := 0.0;           // 零值常量，避免裸字面量 [无量纲] / zero constant, avoids a bare literal [dimensionless]
END_VAR

// 段 0｜输出与错误状态预置 / segment 0, preset outputs and error status
eErr := 0;                                     // 预置无错误 / preset no error
bError := FALSE;                               // 预置无故障 / preset no fault
bOut := FALSE;                                 // 输出先断开，安全侧 / preset the output off, safe side
fDutyApplied := DL_SSR_DUTY_MIN;               // 生效占空先归零 / preset the duty to zero
tOnTime := T#0MS;                              // 导通时长先归零 / preset the conducted time to zero

// 段 1｜周期参数闸：周期非法时宁可断热，绝不满功率长通 / segment 1, period gate, a wrong period must never mean full power
IF (tCycleTime < DL_SSR_CYCLE_MIN) OR (tCycleTime > DL_SSR_CYCLE_MAX) THEN
    eErr := 16#0003_032D;                      // 周期非法故障码 / illegal period fault id
    bError := TRUE;                            // 置故障标志 / raise the error flag
    bOut := FALSE;                             // 输出强制断开 / force the output off
    fDutyApplied := DL_SSR_DUTY_MIN;           // 生效占空归零 / effective duty to zero
    tOnTime := T#0MS;                          // 导通时长为 0 / conducted time zero
    bLoadOpen := bLoadLatch;                   // 锁存状态照常回读 / the latch stays readable
    RETURN;                                    // 故障级提前返回 / early return on fault
END_IF

// 段 2｜占空与诊断参数闸：双侧钳位并置信息码 / segment 2, duty and diagnostic parameter gates
fDutyEff := MIN(MAX(fPowerDemand, DL_SSR_DUTY_MIN), DL_SSR_DUTY_MAX); // 占空双侧钳位 / clamp the duty both sides
IF ABS(fDutyEff - fPowerDemand) > DL_FLOAT_EPS THEN
    eErr := 16#0003_0168;                      // 占空钳位提示（信息级不置故障）/ duty clamp hint, info level never raises a fault
END_IF
fMinDutyEff := MIN(MAX(fMinDutyForCurrent, DL_SSR_MIND_MIN), DL_SSR_MIND_MAX); // 电流判定占空双侧钳位 / clamp the current duty threshold both sides
tWindowEff := MIN(MAX(tCurrentWindow, DL_SSR_WIN_MIN), DL_SSR_WIN_MAX);        // 确认窗双侧钳位 / clamp the confirmation window both sides

// 段 3｜边沿实例无条件周期刷新（红线：严禁放入条件分支）/ segment 3, unconditional edge refresh
fbTrigReset(CLK := bReset);
fbTrigSync(CLK := bSyncPulse);
IF fbTrigSync.Q THEN
    bForceRestart := TRUE;                     // 同步脉冲到来，本拍强制重启周期相位 / a sync pulse forces a phase restart this cycle
END_IF

// 段 4｜周期相位与电流缺失两个定时器无条件调用 / segment 4, unconditional calls of the phase and current timers
bCycleHold := (NOT fbCycle.Q) AND (NOT bForceRestart); // 自复位逻辑：定时器到期或强制重启即掉一拍 IN / self-reset logic, the input drops for one cycle on expiry or forced restart
fbCycle(IN := bEnable AND bCycleHold, PT := tCycleTime); // 周期相位定时器 / cycle phase timer
fCycleMs := TIME_TO_REAL(tCycleTime);          // 周期毫秒值 / cycle in milliseconds
fOnMs := fDutyEff / DL_SSR_PCT_SCALE * fCycleMs; // 应导通毫秒数 / target conducted milliseconds
tOnTarget := REAL_TO_TIME(fOnMs);               // 转 TIME 后与 ET 直接比较，不转 REAL / converted to TIME so it compares with ET without any REAL conversion
bForceRestart := FALSE;                        // 强制重启标志用后即清 / the forced restart flag is consumed and cleared
fbNoCurrent(IN := bEnable AND (fDutyEff >= fMinDutyEff) AND (NOT bCurrentFeedback) AND (NOT bLoadLatch), PT := tWindowEff); // 电流缺失确认定时器 / current absence confirmation timer

// 段 5｜占空镜像（输出已在段 0 预置为断开）/ segment 5, publish the duty, the output was already preset off in segment zero
fDutyApplied := fDutyEff;                      // 占空镜像 / publish the duty

// 段 6｜复位沿清断线锁存（优先于诊断）/ segment 6, reset clears the open circuit latch
IF fbTrigReset.Q THEN
    bLoadLatch := FALSE;                       // 清锁存 / clear the latch
END_IF

// 段 7｜断线诊断：占空足量却无电流超确认窗，即锁存开路 / segment 7, open circuit diagnosis
IF fbNoCurrent.Q THEN
    bLoadLatch := TRUE;                        // 锁存开路 / latch the open circuit
    eErr := 16#0003_032E;                      // 回路开路故障码 / open circuit fault id
    bError := TRUE;                            // 置故障标志 / raise the error flag
END_IF

// 段 8｜PWM 通断判定：零占空不启监视，占空已达导通阈值才允许导通 / segment 8, PWM conduction decision
IF (NOT bEnable) OR bLoadLatch THEN
    bOut := FALSE;                             // 失能或锁存故障一律断输出 / disabled or latched fault forces the output off
    tOnTime := T#0MS;                          // 导通时长归零 / conducted time zero
ELSIF fDutyEff < DL_SSR_ON_EPS THEN
    bOut := FALSE;                             // 占空低于导通阈值，强制全断（信息级提示）/ duty below the threshold forces a full off, info level hint
    tOnTime := T#0MS;                          // 导通时长归零 / conducted time zero
    eErr := 16#0003_0168;                      // 零占空提示（信息级不置故障）/ zero duty hint, info level never raises a fault
ELSIF fDutyEff >= DL_SSR_DUTY_MAX THEN
    bOut := TRUE;                              // 满占空长通 / full duty keeps the output on
    tOnTime := fbCycle.ET;                     // 导通时长取相位 / conducted time follows the phase
ELSE
    IF fbCycle.ET < tOnTarget THEN
        bOut := TRUE;                          // 相位未到导通目标，保持导通 / the phase is below the on target, keep conducting
    ELSE
        bOut := FALSE;                         // 相位越过导通目标，断开 / the phase passed the on target, switch off
    END_IF
    tOnTime := fbCycle.ET;                     // 导通时长取相位 / conducted time follows the phase
END_IF

// 段 9｜锁存对外输出 / segment 9, publish the latch
bLoadOpen := bLoadLatch;                       // 回路开路输出 / open circuit output
END_FUNCTION_BLOCK
